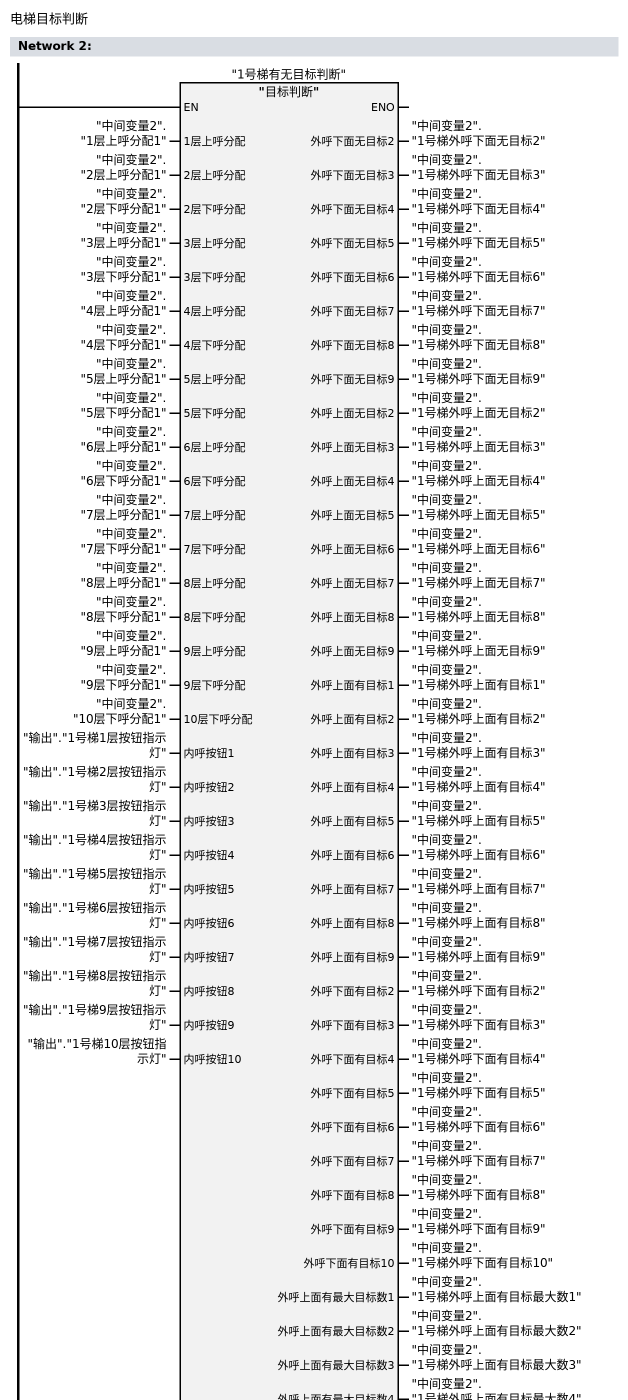
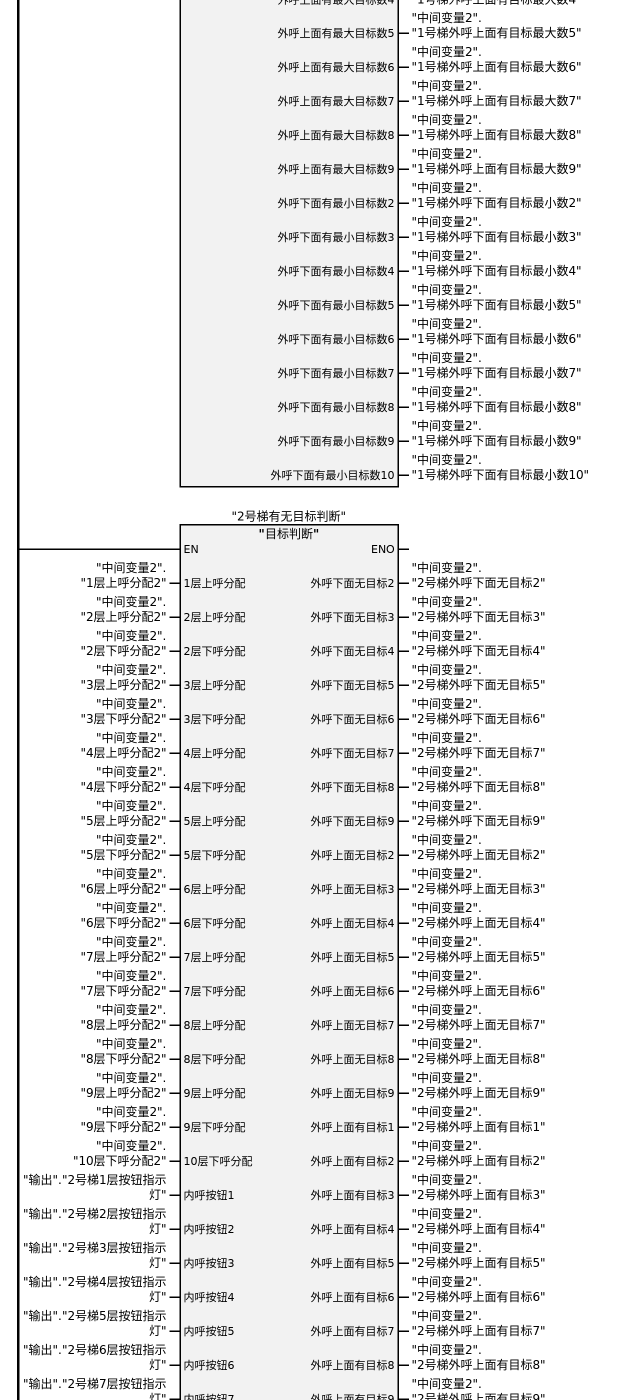
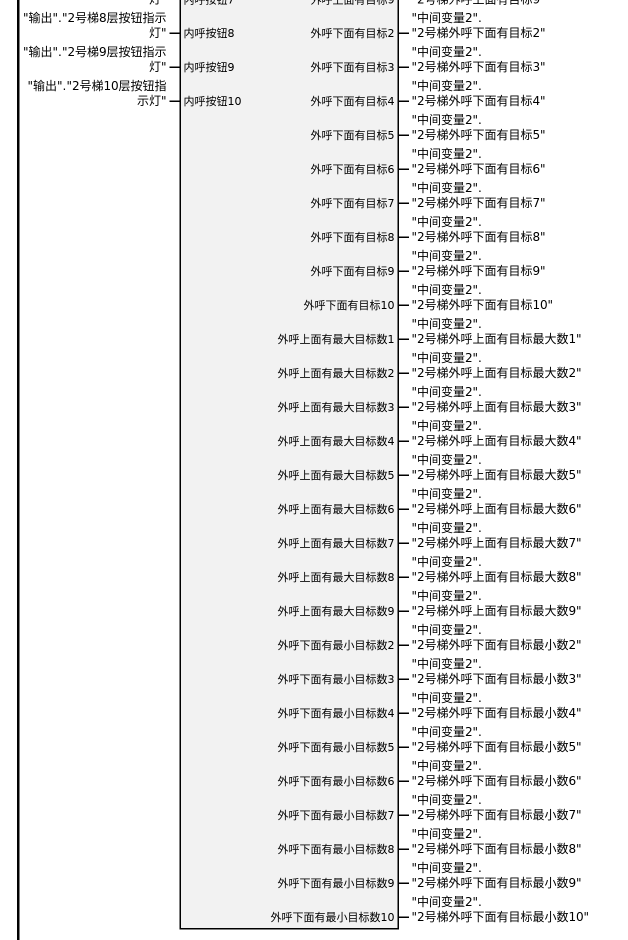
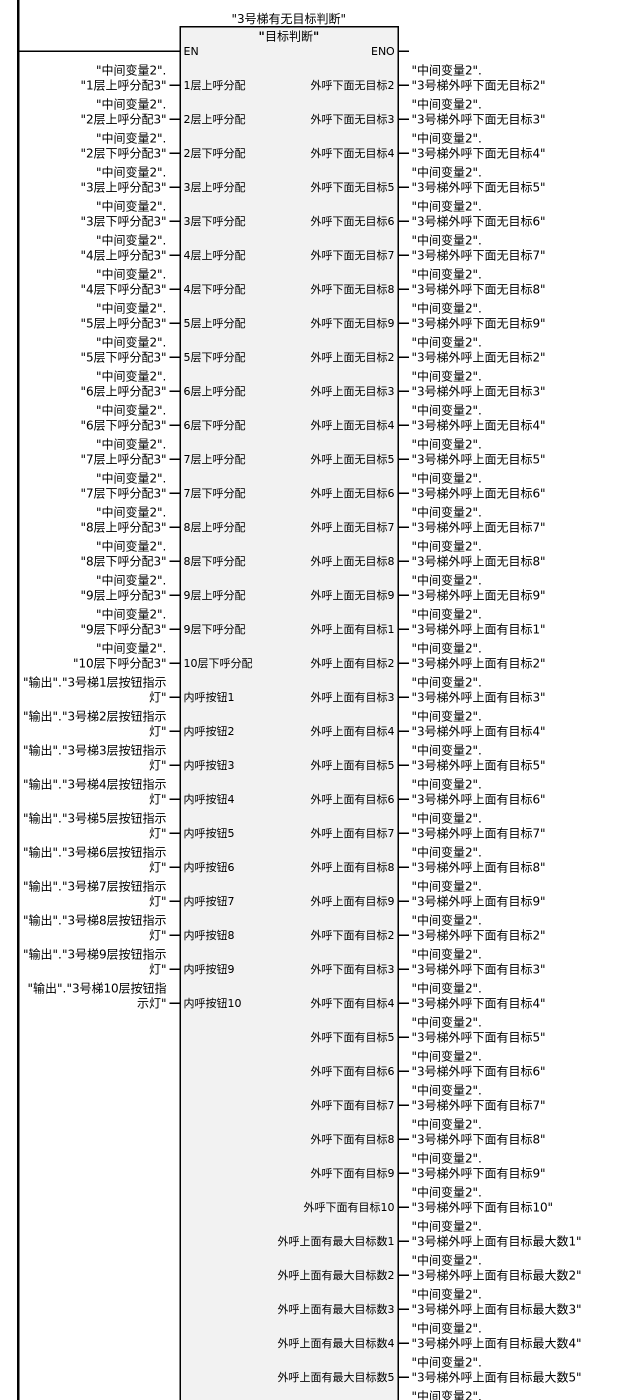
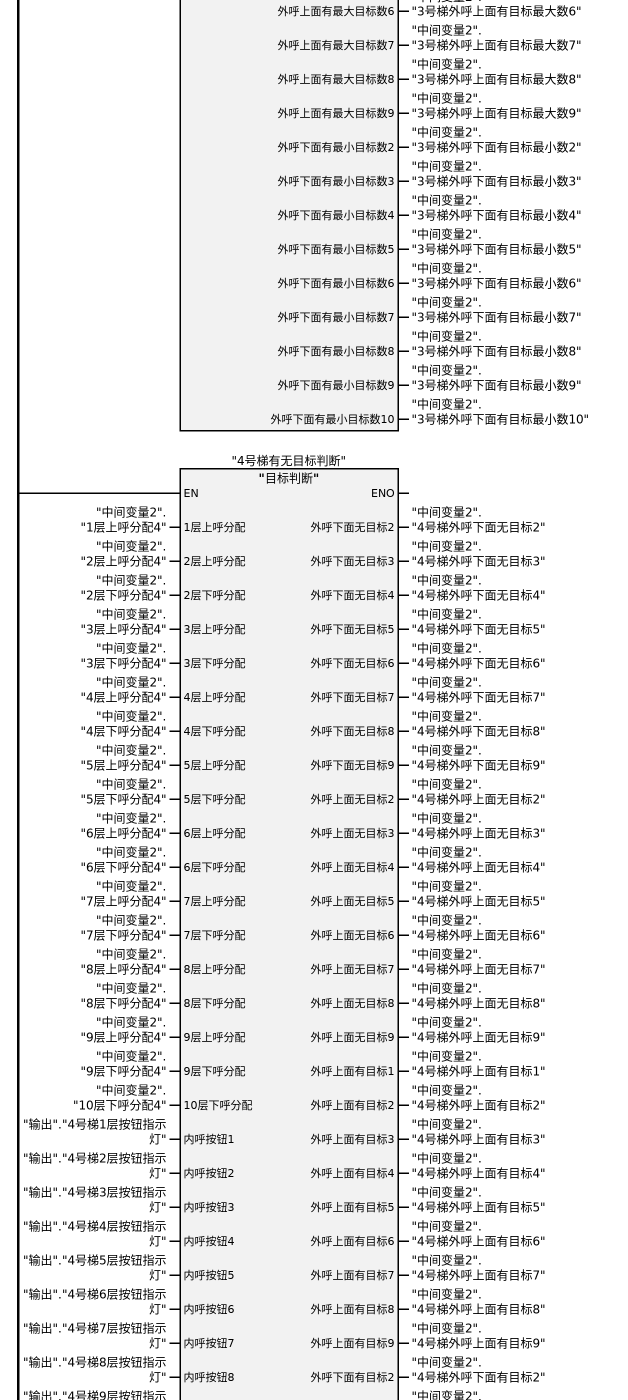
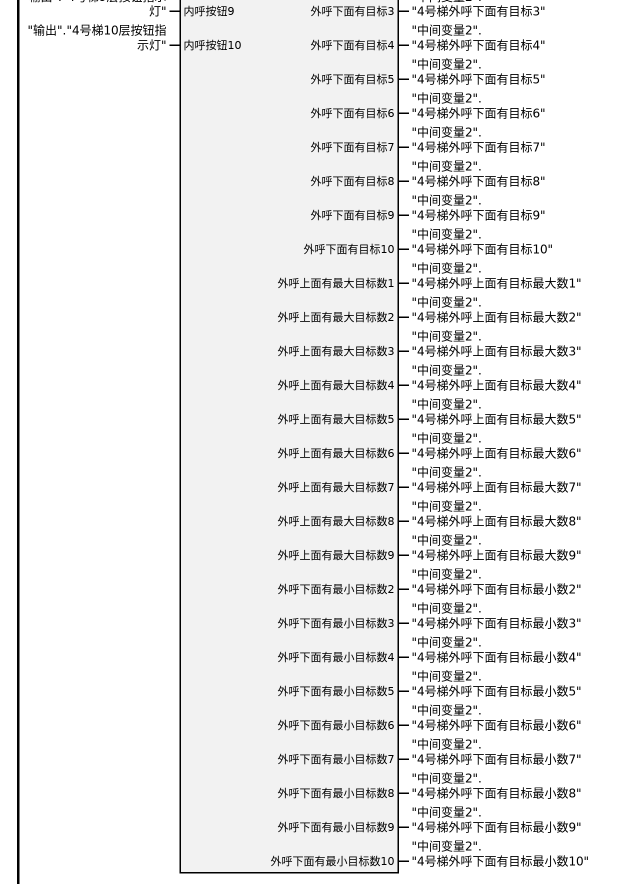
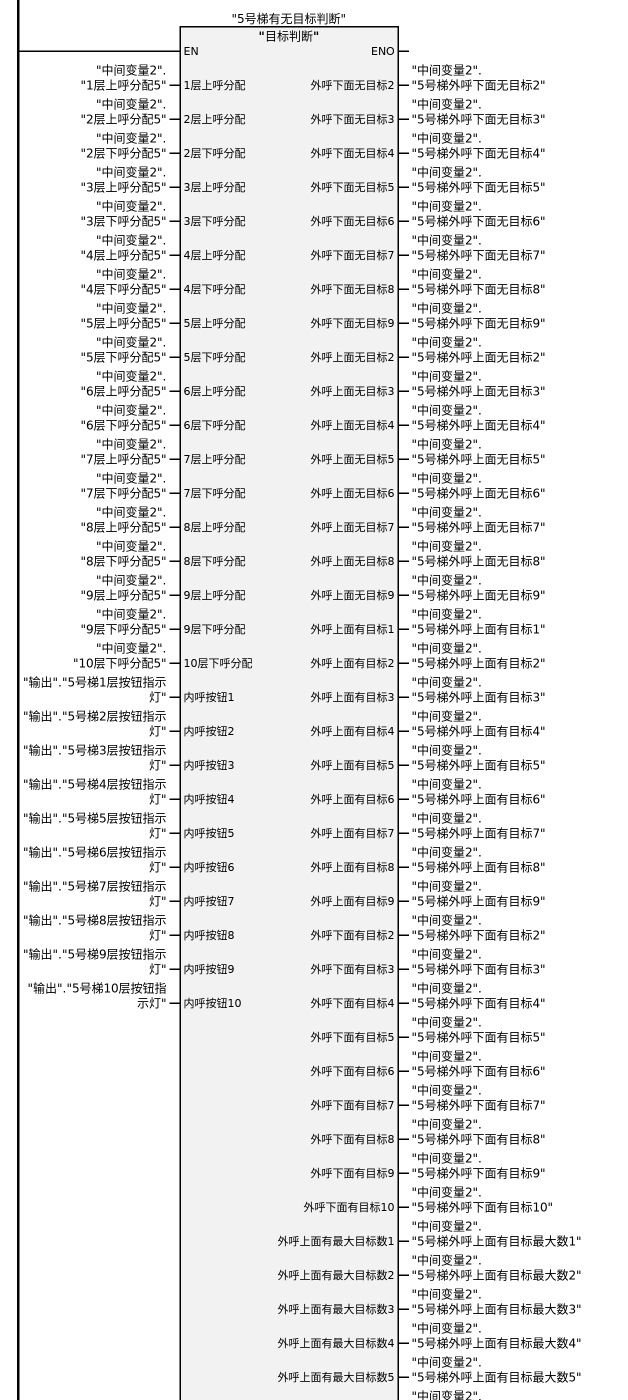
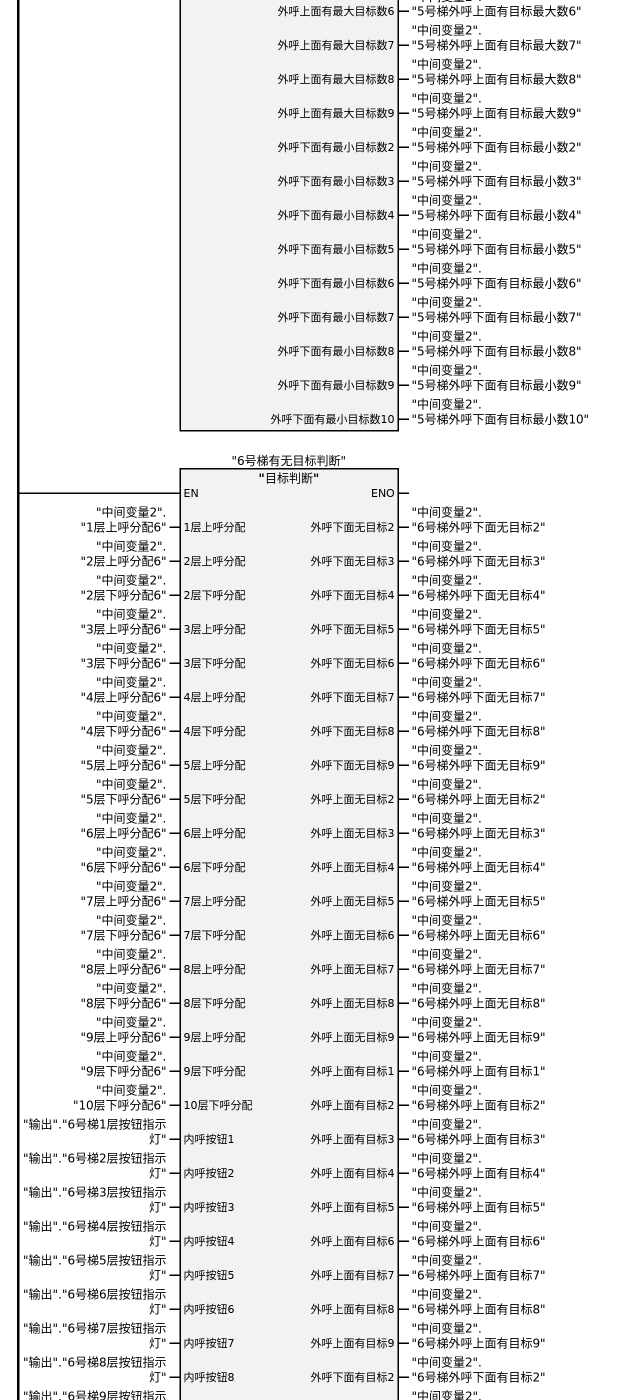
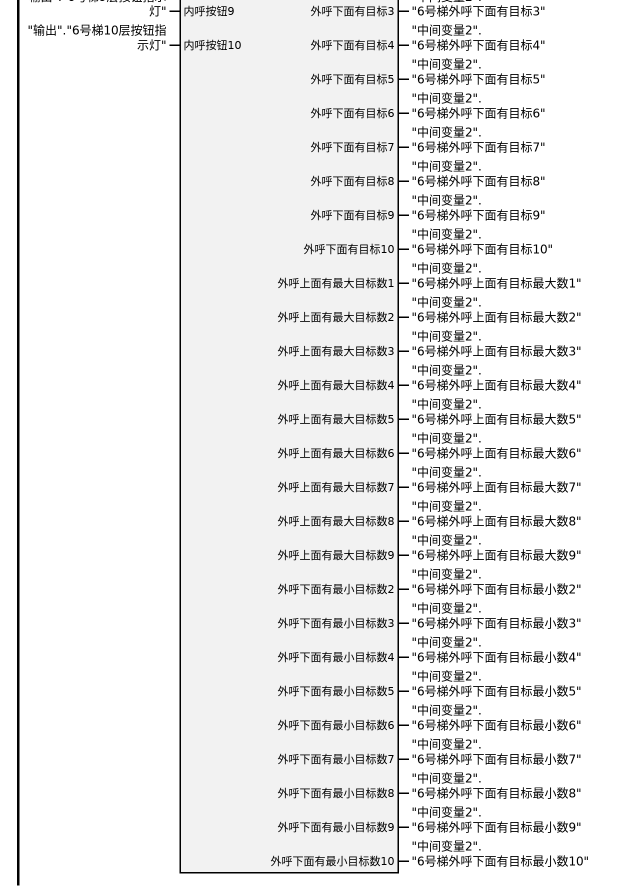
   RUNG wire#powerrail
      "1号梯有无目标判断"("1层上呼分配" := "中间变量2"."1层上呼分配1", "2层上呼分配" := "中间变量2"."2层上呼分配1", "2层下呼分配" := "中间变量2"."2层下呼分配1", "3层上呼分配" := "中间变量2"."3层上呼分配1", "3层下呼分配" := "中间变量2"."3层下呼分配1", "4层上呼分配" := "中间变量2"."4层上呼分配1", "4层下呼分配" := "中间变量2"."4层下呼分配1", "5层上呼分配" := "中间变量2"."5层上呼分配1", "5层下呼分配" := "中间变量2"."5层下呼分配1", "6层上呼分配" := "中间变量2"."6层上呼分配1", "6层下呼分配" := "中间变量2"."6层下呼分配1", "7层上呼分配" := "中间变量2"."7层上呼分配1", "7层下呼分配" := "中间变量2"."7层下呼分配1", "8层上呼分配" := "中间变量2"."8层上呼分配1", "8层下呼分配" := "中间变量2"."8层下呼分配1", "9层上呼分配" := "中间变量2"."9层上呼分配1", "9层下呼分配" := "中间变量2"."9层下呼分配1", "10层下呼分配" := "中间变量2"."10层下呼分配1", 内呼按钮1 := "输出"."1号梯1层按钮指示灯", 内呼按钮2 := "输出"."1号梯2层按钮指示灯", 内呼按钮3 := "输出"."1号梯3层按钮指示灯", 内呼按钮4 := "输出"."1号梯4层按钮指示灯", 内呼按钮5 := "输出"."1号梯5层按钮指示灯", 内呼按钮6 := "输出"."1号梯6层按钮指示灯", 内呼按钮7 := "输出"."1号梯7层按钮指示灯", 内呼按钮8 := "输出"."1号梯8层按钮指示灯", 内呼按钮9 := "输出"."1号梯9层按钮指示灯", 内呼按钮10 := "输出"."1号梯10层按钮指示灯", 外呼下面无目标2 => "中间变量2"."1号梯外呼下面无目标2", 外呼下面无目标3 => "中间变量2"."1号梯外呼下面无目标3", 外呼下面无目标4 => "中间变量2"."1号梯外呼下面无目标4", 外呼下面无目标5 => "中间变量2"."1号梯外呼下面无目标5", 外呼下面无目标6 => "中间变量2"."1号梯外呼下面无目标6", 外呼下面无目标7 => "中间变量2"."1号梯外呼下面无目标7", 外呼下面无目标8 => "中间变量2"."1号梯外呼下面无目标8", 外呼下面无目标9 => "中间变量2"."1号梯外呼下面无目标9", 外呼上面无目标2 => "中间变量2"."1号梯外呼上面无目标2", 外呼上面无目标3 => "中间变量2"."1号梯外呼上面无目标3", 外呼上面无目标4 => "中间变量2"."1号梯外呼上面无目标4", 外呼上面无目标5 => "中间变量2"."1号梯外呼上面无目标5", 外呼上面无目标6 => "中间变量2"."1号梯外呼上面无目标6", 外呼上面无目标7 => "中间变量2"."1号梯外呼上面无目标7", 外呼上面无目标8 => "中间变量2"."1号梯外呼上面无目标8", 外呼上面无目标9 => "中间变量2"."1号梯外呼上面无目标9", 外呼上面有目标1 => "中间变量2"."1号梯外呼上面有目标1", 外呼上面有目标2 => "中间变量2"."1号梯外呼上面有目标2", 外呼上面有目标3 => "中间变量2"."1号梯外呼上面有目标3", 外呼上面有目标4 => "中间变量2"."1号梯外呼上面有目标4", 外呼上面有目标5 => "中间变量2"."1号梯外呼上面有目标5", 外呼上面有目标6 => "中间变量2"."1号梯外呼上面有目标6", 外呼上面有目标7 => "中间变量2"."1号梯外呼上面有目标7", 外呼上面有目标8 => "中间变量2"."1号梯外呼上面有目标8", 外呼上面有目标9 => "中间变量2"."1号梯外呼上面有目标9", 外呼下面有目标2 => "中间变量2"."1号梯外呼下面有目标2", 外呼下面有目标3 => "中间变量2"."1号梯外呼下面有目标3", 外呼下面有目标4 => "中间变量2"."1号梯外呼下面有目标4", 外呼下面有目标5 => "中间变量2"."1号梯外呼下面有目标5", 外呼下面有目标6 => "中间变量2"."1号梯外呼下面有目标6", 外呼下面有目标7 => "中间变量2"."1号梯外呼下面有目标7", 外呼下面有目标8 => "中间变量2"."1号梯外呼下面有目标8", 外呼下面有目标9 => "中间变量2"."1号梯外呼下面有目标9", 外呼下面有目标10 => "中间变量2"."1号梯外呼下面有目标10", 外呼上面有最大目标数1 => "中间变量2"."1号梯外呼上面有目标最大数1", 外呼上面有最大目标数2 => "中间变量2"."1号梯外呼上面有目标最大数2", 外呼上面有最大目标数3 => "中间变量2"."1号梯外呼上面有目标最大数3", 外呼上面有最大目标数4 => "中间变量2"."1号梯外呼上面有目标最大数4", 外呼上面有最大目标数5 => "中间变量2"."1号梯外呼上面有目标最大数5", 外呼上面有最大目标数6 => "中间变量2"."1号梯外呼上面有目标最大数6", 外呼上面有最大目标数7 => "中间变量2"."1号梯外呼上面有目标最大数7", 外呼上面有最大目标数8 => "中间变量2"."1号梯外呼上面有目标最大数8", 外呼上面有最大目标数9 => "中间变量2"."1号梯外呼上面有目标最大数9", 外呼下面有最小目标数2 => "中间变量2"."1号梯外呼下面有目标最小数2", 外呼下面有最小目标数3 => "中间变量2"."1号梯外呼下面有目标最小数3", 外呼下面有最小目标数4 => "中间变量2"."1号梯外呼下面有目标最小数4", 外呼下面有最小目标数5 => "中间变量2"."1号梯外呼下面有目标最小数5", 外呼下面有最小目标数6 => "中间变量2"."1号梯外呼下面有目标最小数6", 外呼下面有最小目标数7 => "中间变量2"."1号梯外呼下面有目标最小数7", 外呼下面有最小目标数8 => "中间变量2"."1号梯外呼下面有目标最小数8", 外呼下面有最小目标数9 => "中间变量2"."1号梯外呼下面有目标最小数9", 外呼下面有最小目标数10 => "中间变量2"."1号梯外呼下面有目标最小数10")
   END_RUNG
   RUNG wire#powerrail
      "2号梯有无目标判断"("1层上呼分配" := "中间变量2"."1层上呼分配2", "2层上呼分配" := "中间变量2"."2层上呼分配2", "2层下呼分配" := "中间变量2"."2层下呼分配2", "3层上呼分配" := "中间变量2"."3层上呼分配2", "3层下呼分配" := "中间变量2"."3层下呼分配2", "4层上呼分配" := "中间变量2"."4层上呼分配2", "4层下呼分配" := "中间变量2"."4层下呼分配2", "5层上呼分配" := "中间变量2"."5层上呼分配2", "5层下呼分配" := "中间变量2"."5层下呼分配2", "6层上呼分配" := "中间变量2"."6层上呼分配2", "6层下呼分配" := "中间变量2"."6层下呼分配2", "7层上呼分配" := "中间变量2"."7层上呼分配2", "7层下呼分配" := "中间变量2"."7层下呼分配2", "8层上呼分配" := "中间变量2"."8层上呼分配2", "8层下呼分配" := "中间变量2"."8层下呼分配2", "9层上呼分配" := "中间变量2"."9层上呼分配2", "9层下呼分配" := "中间变量2"."9层下呼分配2", "10层下呼分配" := "中间变量2"."10层下呼分配2", 内呼按钮1 := "输出"."2号梯1层按钮指示灯", 内呼按钮2 := "输出"."2号梯2层按钮指示灯", 内呼按钮3 := "输出"."2号梯3层按钮指示灯", 内呼按钮4 := "输出"."2号梯4层按钮指示灯", 内呼按钮5 := "输出"."2号梯5层按钮指示灯", 内呼按钮6 := "输出"."2号梯6层按钮指示灯", 内呼按钮7 := "输出"."2号梯7层按钮指示灯", 内呼按钮8 := "输出"."2号梯8层按钮指示灯", 内呼按钮9 := "输出"."2号梯9层按钮指示灯", 内呼按钮10 := "输出"."2号梯10层按钮指示灯", 外呼下面无目标2 => "中间变量2"."2号梯外呼下面无目标2", 外呼下面无目标3 => "中间变量2"."2号梯外呼下面无目标3", 外呼下面无目标4 => "中间变量2"."2号梯外呼下面无目标4", 外呼下面无目标5 => "中间变量2"."2号梯外呼下面无目标5", 外呼下面无目标6 => "中间变量2"."2号梯外呼下面无目标6", 外呼下面无目标7 => "中间变量2"."2号梯外呼下面无目标7", 外呼下面无目标8 => "中间变量2"."2号梯外呼下面无目标8", 外呼下面无目标9 => "中间变量2"."2号梯外呼下面无目标9", 外呼上面无目标2 => "中间变量2"."2号梯外呼上面无目标2", 外呼上面无目标3 => "中间变量2"."2号梯外呼上面无目标3", 外呼上面无目标4 => "中间变量2"."2号梯外呼上面无目标4", 外呼上面无目标5 => "中间变量2"."2号梯外呼上面无目标5", 外呼上面无目标6 => "中间变量2"."2号梯外呼上面无目标6", 外呼上面无目标7 => "中间变量2"."2号梯外呼上面无目标7", 外呼上面无目标8 => "中间变量2"."2号梯外呼上面无目标8", 外呼上面无目标9 => "中间变量2"."2号梯外呼上面无目标9", 外呼上面有目标1 => "中间变量2"."2号梯外呼上面有目标1", 外呼上面有目标2 => "中间变量2"."2号梯外呼上面有目标2", 外呼上面有目标3 => "中间变量2"."2号梯外呼上面有目标3", 外呼上面有目标4 => "中间变量2"."2号梯外呼上面有目标4", 外呼上面有目标5 => "中间变量2"."2号梯外呼上面有目标5", 外呼上面有目标6 => "中间变量2"."2号梯外呼上面有目标6", 外呼上面有目标7 => "中间变量2"."2号梯外呼上面有目标7", 外呼上面有目标8 => "中间变量2"."2号梯外呼上面有目标8", 外呼上面有目标9 => "中间变量2"."2号梯外呼上面有目标9", 外呼下面有目标2 => "中间变量2"."2号梯外呼下面有目标2", 外呼下面有目标3 => "中间变量2"."2号梯外呼下面有目标3", 外呼下面有目标4 => "中间变量2"."2号梯外呼下面有目标4", 外呼下面有目标5 => "中间变量2"."2号梯外呼下面有目标5", 外呼下面有目标6 => "中间变量2"."2号梯外呼下面有目标6", 外呼下面有目标7 => "中间变量2"."2号梯外呼下面有目标7", 外呼下面有目标8 => "中间变量2"."2号梯外呼下面有目标8", 外呼下面有目标9 => "中间变量2"."2号梯外呼下面有目标9", 外呼下面有目标10 => "中间变量2"."2号梯外呼下面有目标10", 外呼上面有最大目标数1 => "中间变量2"."2号梯外呼上面有目标最大数1", 外呼上面有最大目标数2 => "中间变量2"."2号梯外呼上面有目标最大数2", 外呼上面有最大目标数3 => "中间变量2"."2号梯外呼上面有目标最大数3", 外呼上面有最大目标数4 => "中间变量2"."2号梯外呼上面有目标最大数4", 外呼上面有最大目标数5 => "中间变量2"."2号梯外呼上面有目标最大数5", 外呼上面有最大目标数6 => "中间变量2"."2号梯外呼上面有目标最大数6", 外呼上面有最大目标数7 => "中间变量2"."2号梯外呼上面有目标最大数7", 外呼上面有最大目标数8 => "中间变量2"."2号梯外呼上面有目标最大数8", 外呼上面有最大目标数9 => "中间变量2"."2号梯外呼上面有目标最大数9", 外呼下面有最小目标数2 => "中间变量2"."2号梯外呼下面有目标最小数2", 外呼下面有最小目标数3 => "中间变量2"."2号梯外呼下面有目标最小数3", 外呼下面有最小目标数4 => "中间变量2"."2号梯外呼下面有目标最小数4", 外呼下面有最小目标数5 => "中间变量2"."2号梯外呼下面有目标最小数5", 外呼下面有最小目标数6 => "中间变量2"."2号梯外呼下面有目标最小数6", 外呼下面有最小目标数7 => "中间变量2"."2号梯外呼下面有目标最小数7", 外呼下面有最小目标数8 => "中间变量2"."2号梯外呼下面有目标最小数8", 外呼下面有最小目标数9 => "中间变量2"."2号梯外呼下面有目标最小数9", 外呼下面有最小目标数10 => "中间变量2"."2号梯外呼下面有目标最小数10")
   END_RUNG
   RUNG wire#powerrail
      "3号梯有无目标判断"("1层上呼分配" := "中间变量2"."1层上呼分配3", "2层上呼分配" := "中间变量2"."2层上呼分配3", "2层下呼分配" := "中间变量2"."2层下呼分配3", "3层上呼分配" := "中间变量2"."3层上呼分配3", "3层下呼分配" := "中间变量2"."3层下呼分配3", "4层上呼分配" := "中间变量2"."4层上呼分配3", "4层下呼分配" := "中间变量2"."4层下呼分配3", "5层上呼分配" := "中间变量2"."5层上呼分配3", "5层下呼分配" := "中间变量2"."5层下呼分配3", "6层上呼分配" := "中间变量2"."6层上呼分配3", "6层下呼分配" := "中间变量2"."6层下呼分配3", "7层上呼分配" := "中间变量2"."7层上呼分配3", "7层下呼分配" := "中间变量2"."7层下呼分配3", "8层上呼分配" := "中间变量2"."8层上呼分配3", "8层下呼分配" := "中间变量2"."8层下呼分配3", "9层上呼分配" := "中间变量2"."9层上呼分配3", "9层下呼分配" := "中间变量2"."9层下呼分配3", "10层下呼分配" := "中间变量2"."10层下呼分配3", 内呼按钮1 := "输出"."3号梯1层按钮指示灯", 内呼按钮2 := "输出"."3号梯2层按钮指示灯", 内呼按钮3 := "输出"."3号梯3层按钮指示灯", 内呼按钮4 := "输出"."3号梯4层按钮指示灯", 内呼按钮5 := "输出"."3号梯5层按钮指示灯", 内呼按钮6 := "输出"."3号梯6层按钮指示灯", 内呼按钮7 := "输出"."3号梯7层按钮指示灯", 内呼按钮8 := "输出"."3号梯8层按钮指示灯", 内呼按钮9 := "输出"."3号梯9层按钮指示灯", 内呼按钮10 := "输出"."3号梯10层按钮指示灯", 外呼下面无目标2 => "中间变量2"."3号梯外呼下面无目标2", 外呼下面无目标3 => "中间变量2"."3号梯外呼下面无目标3", 外呼下面无目标4 => "中间变量2"."3号梯外呼下面无目标4", 外呼下面无目标5 => "中间变量2"."3号梯外呼下面无目标5", 外呼下面无目标6 => "中间变量2"."3号梯外呼下面无目标6", 外呼下面无目标7 => "中间变量2"."3号梯外呼下面无目标7", 外呼下面无目标8 => "中间变量2"."3号梯外呼下面无目标8", 外呼下面无目标9 => "中间变量2"."3号梯外呼下面无目标9", 外呼上面无目标2 => "中间变量2"."3号梯外呼上面无目标2", 外呼上面无目标3 => "中间变量2"."3号梯外呼上面无目标3", 外呼上面无目标4 => "中间变量2"."3号梯外呼上面无目标4", 外呼上面无目标5 => "中间变量2"."3号梯外呼上面无目标5", 外呼上面无目标6 => "中间变量2"."3号梯外呼上面无目标6", 外呼上面无目标7 => "中间变量2"."3号梯外呼上面无目标7", 外呼上面无目标8 => "中间变量2"."3号梯外呼上面无目标8", 外呼上面无目标9 => "中间变量2"."3号梯外呼上面无目标9", 外呼上面有目标1 => "中间变量2"."3号梯外呼上面有目标1", 外呼上面有目标2 => "中间变量2"."3号梯外呼上面有目标2", 外呼上面有目标3 => "中间变量2"."3号梯外呼上面有目标3", 外呼上面有目标4 => "中间变量2"."3号梯外呼上面有目标4", 外呼上面有目标5 => "中间变量2"."3号梯外呼上面有目标5", 外呼上面有目标6 => "中间变量2"."3号梯外呼上面有目标6", 外呼上面有目标7 => "中间变量2"."3号梯外呼上面有目标7", 外呼上面有目标8 => "中间变量2"."3号梯外呼上面有目标8", 外呼上面有目标9 => "中间变量2"."3号梯外呼上面有目标9", 外呼下面有目标2 => "中间变量2"."3号梯外呼下面有目标2", 外呼下面有目标3 => "中间变量2"."3号梯外呼下面有目标3", 外呼下面有目标4 => "中间变量2"."3号梯外呼下面有目标4", 外呼下面有目标5 => "中间变量2"."3号梯外呼下面有目标5", 外呼下面有目标6 => "中间变量2"."3号梯外呼下面有目标6", 外呼下面有目标7 => "中间变量2"."3号梯外呼下面有目标7", 外呼下面有目标8 => "中间变量2"."3号梯外呼下面有目标8", 外呼下面有目标9 => "中间变量2"."3号梯外呼下面有目标9", 外呼下面有目标10 => "中间变量2"."3号梯外呼下面有目标10", 外呼上面有最大目标数1 => "中间变量2"."3号梯外呼上面有目标最大数1", 外呼上面有最大目标数2 => "中间变量2"."3号梯外呼上面有目标最大数2", 外呼上面有最大目标数3 => "中间变量2"."3号梯外呼上面有目标最大数3", 外呼上面有最大目标数4 => "中间变量2"."3号梯外呼上面有目标最大数4", 外呼上面有最大目标数5 => "中间变量2"."3号梯外呼上面有目标最大数5", 外呼上面有最大目标数6 => "中间变量2"."3号梯外呼上面有目标最大数6", 外呼上面有最大目标数7 => "中间变量2"."3号梯外呼上面有目标最大数7", 外呼上面有最大目标数8 => "中间变量2"."3号梯外呼上面有目标最大数8", 外呼上面有最大目标数9 => "中间变量2"."3号梯外呼上面有目标最大数9", 外呼下面有最小目标数2 => "中间变量2"."3号梯外呼下面有目标最小数2", 外呼下面有最小目标数3 => "中间变量2"."3号梯外呼下面有目标最小数3", 外呼下面有最小目标数4 => "中间变量2"."3号梯外呼下面有目标最小数4", 外呼下面有最小目标数5 => "中间变量2"."3号梯外呼下面有目标最小数5", 外呼下面有最小目标数6 => "中间变量2"."3号梯外呼下面有目标最小数6", 外呼下面有最小目标数7 => "中间变量2"."3号梯外呼下面有目标最小数7", 外呼下面有最小目标数8 => "中间变量2"."3号梯外呼下面有目标最小数8", 外呼下面有最小目标数9 => "中间变量2"."3号梯外呼下面有目标最小数9", 外呼下面有最小目标数10 => "中间变量2"."3号梯外呼下面有目标最小数10")
   END_RUNG
   RUNG wire#powerrail
      "4号梯有无目标判断"("1层上呼分配" := "中间变量2"."1层上呼分配4", "2层上呼分配" := "中间变量2"."2层上呼分配4", "2层下呼分配" := "中间变量2"."2层下呼分配4", "3层上呼分配" := "中间变量2"."3层上呼分配4", "3层下呼分配" := "中间变量2"."3层下呼分配4", "4层上呼分配" := "中间变量2"."4层上呼分配4", "4层下呼分配" := "中间变量2"."4层下呼分配4", "5层上呼分配" := "中间变量2"."5层上呼分配4", "5层下呼分配" := "中间变量2"."5层下呼分配4", "6层上呼分配" := "中间变量2"."6层上呼分配4", "6层下呼分配" := "中间变量2"."6层下呼分配4", "7层上呼分配" := "中间变量2"."7层上呼分配4", "7层下呼分配" := "中间变量2"."7层下呼分配4", "8层上呼分配" := "中间变量2"."8层上呼分配4", "8层下呼分配" := "中间变量2"."8层下呼分配4", "9层上呼分配" := "中间变量2"."9层上呼分配4", "9层下呼分配" := "中间变量2"."9层下呼分配4", "10层下呼分配" := "中间变量2"."10层下呼分配4", 内呼按钮1 := "输出"."4号梯1层按钮指示灯", 内呼按钮2 := "输出"."4号梯2层按钮指示灯", 内呼按钮3 := "输出"."4号梯3层按钮指示灯", 内呼按钮4 := "输出"."4号梯4层按钮指示灯", 内呼按钮5 := "输出"."4号梯5层按钮指示灯", 内呼按钮6 := "输出"."4号梯6层按钮指示灯", 内呼按钮7 := "输出"."4号梯7层按钮指示灯", 内呼按钮8 := "输出"."4号梯8层按钮指示灯", 内呼按钮9 := "输出"."4号梯9层按钮指示灯", 内呼按钮10 := "输出"."4号梯10层按钮指示灯", 外呼下面无目标2 => "中间变量2"."4号梯外呼下面无目标2", 外呼下面无目标3 => "中间变量2"."4号梯外呼下面无目标3", 外呼下面无目标4 => "中间变量2"."4号梯外呼下面无目标4", 外呼下面无目标5 => "中间变量2"."4号梯外呼下面无目标5", 外呼下面无目标6 => "中间变量2"."4号梯外呼下面无目标6", 外呼下面无目标7 => "中间变量2"."4号梯外呼下面无目标7", 外呼下面无目标8 => "中间变量2"."4号梯外呼下面无目标8", 外呼下面无目标9 => "中间变量2"."4号梯外呼下面无目标9", 外呼上面无目标2 => "中间变量2"."4号梯外呼上面无目标2", 外呼上面无目标3 => "中间变量2"."4号梯外呼上面无目标3", 外呼上面无目标4 => "中间变量2"."4号梯外呼上面无目标4", 外呼上面无目标5 => "中间变量2"."4号梯外呼上面无目标5", 外呼上面无目标6 => "中间变量2"."4号梯外呼上面无目标6", 外呼上面无目标7 => "中间变量2"."4号梯外呼上面无目标7", 外呼上面无目标8 => "中间变量2"."4号梯外呼上面无目标8", 外呼上面无目标9 => "中间变量2"."4号梯外呼上面无目标9", 外呼上面有目标1 => "中间变量2"."4号梯外呼上面有目标1", 外呼上面有目标2 => "中间变量2"."4号梯外呼上面有目标2", 外呼上面有目标3 => "中间变量2"."4号梯外呼上面有目标3", 外呼上面有目标4 => "中间变量2"."4号梯外呼上面有目标4", 外呼上面有目标5 => "中间变量2"."4号梯外呼上面有目标5", 外呼上面有目标6 => "中间变量2"."4号梯外呼上面有目标6", 外呼上面有目标7 => "中间变量2"."4号梯外呼上面有目标7", 外呼上面有目标8 => "中间变量2"."4号梯外呼上面有目标8", 外呼上面有目标9 => "中间变量2"."4号梯外呼上面有目标9", 外呼下面有目标2 => "中间变量2"."4号梯外呼下面有目标2", 外呼下面有目标3 => "中间变量2"."4号梯外呼下面有目标3", 外呼下面有目标4 => "中间变量2"."4号梯外呼下面有目标4", 外呼下面有目标5 => "中间变量2"."4号梯外呼下面有目标5", 外呼下面有目标6 => "中间变量2"."4号梯外呼下面有目标6", 外呼下面有目标7 => "中间变量2"."4号梯外呼下面有目标7", 外呼下面有目标8 => "中间变量2"."4号梯外呼下面有目标8", 外呼下面有目标9 => "中间变量2"."4号梯外呼下面有目标9", 外呼下面有目标10 => "中间变量2"."4号梯外呼下面有目标10", 外呼上面有最大目标数1 => "中间变量2"."4号梯外呼上面有目标最大数1", 外呼上面有最大目标数2 => "中间变量2"."4号梯外呼上面有目标最大数2", 外呼上面有最大目标数3 => "中间变量2"."4号梯外呼上面有目标最大数3", 外呼上面有最大目标数4 => "中间变量2"."4号梯外呼上面有目标最大数4", 外呼上面有最大目标数5 => "中间变量2"."4号梯外呼上面有目标最大数5", 外呼上面有最大目标数6 => "中间变量2"."4号梯外呼上面有目标最大数6", 外呼上面有最大目标数7 => "中间变量2"."4号梯外呼上面有目标最大数7", 外呼上面有最大目标数8 => "中间变量2"."4号梯外呼上面有目标最大数8", 外呼上面有最大目标数9 => "中间变量2"."4号梯外呼上面有目标最大数9", 外呼下面有最小目标数2 => "中间变量2"."4号梯外呼下面有目标最小数2", 外呼下面有最小目标数3 => "中间变量2"."4号梯外呼下面有目标最小数3", 外呼下面有最小目标数4 => "中间变量2"."4号梯外呼下面有目标最小数4", 外呼下面有最小目标数5 => "中间变量2"."4号梯外呼下面有目标最小数5", 外呼下面有最小目标数6 => "中间变量2"."4号梯外呼下面有目标最小数6", 外呼下面有最小目标数7 => "中间变量2"."4号梯外呼下面有目标最小数7", 外呼下面有最小目标数8 => "中间变量2"."4号梯外呼下面有目标最小数8", 外呼下面有最小目标数9 => "中间变量2"."4号梯外呼下面有目标最小数9", 外呼下面有最小目标数10 => "中间变量2"."4号梯外呼下面有目标最小数10")
   END_RUNG
   RUNG wire#powerrail
      "5号梯有无目标判断"("1层上呼分配" := "中间变量2"."1层上呼分配5", "2层上呼分配" := "中间变量2"."2层上呼分配5", "2层下呼分配" := "中间变量2"."2层下呼分配5", "3层上呼分配" := "中间变量2"."3层上呼分配5", "3层下呼分配" := "中间变量2"."3层下呼分配5", "4层上呼分配" := "中间变量2"."4层上呼分配5", "4层下呼分配" := "中间变量2"."4层下呼分配5", "5层上呼分配" := "中间变量2"."5层上呼分配5", "5层下呼分配" := "中间变量2"."5层下呼分配5", "6层上呼分配" := "中间变量2"."6层上呼分配5", "6层下呼分配" := "中间变量2"."6层下呼分配5", "7层上呼分配" := "中间变量2"."7层上呼分配5", "7层下呼分配" := "中间变量2"."7层下呼分配5", "8层上呼分配" := "中间变量2"."8层上呼分配5", "8层下呼分配" := "中间变量2"."8层下呼分配5", "9层上呼分配" := "中间变量2"."9层上呼分配5", "9层下呼分配" := "中间变量2"."9层下呼分配5", "10层下呼分配" := "中间变量2"."10层下呼分配5", 内呼按钮1 := "输出"."5号梯1层按钮指示灯", 内呼按钮2 := "输出"."5号梯2层按钮指示灯", 内呼按钮3 := "输出"."5号梯3层按钮指示灯", 内呼按钮4 := "输出"."5号梯4层按钮指示灯", 内呼按钮5 := "输出"."5号梯5层按钮指示灯", 内呼按钮6 := "输出"."5号梯6层按钮指示灯", 内呼按钮7 := "输出"."5号梯7层按钮指示灯", 内呼按钮8 := "输出"."5号梯8层按钮指示灯", 内呼按钮9 := "输出"."5号梯9层按钮指示灯", 内呼按钮10 := "输出"."5号梯10层按钮指示灯", 外呼下面无目标2 => "中间变量2"."5号梯外呼下面无目标2", 外呼下面无目标3 => "中间变量2"."5号梯外呼下面无目标3", 外呼下面无目标4 => "中间变量2"."5号梯外呼下面无目标4", 外呼下面无目标5 => "中间变量2"."5号梯外呼下面无目标5", 外呼下面无目标6 => "中间变量2"."5号梯外呼下面无目标6", 外呼下面无目标7 => "中间变量2"."5号梯外呼下面无目标7", 外呼下面无目标8 => "中间变量2"."5号梯外呼下面无目标8", 外呼下面无目标9 => "中间变量2"."5号梯外呼下面无目标9", 外呼上面无目标2 => "中间变量2"."5号梯外呼上面无目标2", 外呼上面无目标3 => "中间变量2"."5号梯外呼上面无目标3", 外呼上面无目标4 => "中间变量2"."5号梯外呼上面无目标4", 外呼上面无目标5 => "中间变量2"."5号梯外呼上面无目标5", 外呼上面无目标6 => "中间变量2"."5号梯外呼上面无目标6", 外呼上面无目标7 => "中间变量2"."5号梯外呼上面无目标7", 外呼上面无目标8 => "中间变量2"."5号梯外呼上面无目标8", 外呼上面无目标9 => "中间变量2"."5号梯外呼上面无目标9", 外呼上面有目标1 => "中间变量2"."5号梯外呼上面有目标1", 外呼上面有目标2 => "中间变量2"."5号梯外呼上面有目标2", 外呼上面有目标3 => "中间变量2"."5号梯外呼上面有目标3", 外呼上面有目标4 => "中间变量2"."5号梯外呼上面有目标4", 外呼上面有目标5 => "中间变量2"."5号梯外呼上面有目标5", 外呼上面有目标6 => "中间变量2"."5号梯外呼上面有目标6", 外呼上面有目标7 => "中间变量2"."5号梯外呼上面有目标7", 外呼上面有目标8 => "中间变量2"."5号梯外呼上面有目标8", 外呼上面有目标9 => "中间变量2"."5号梯外呼上面有目标9", 外呼下面有目标2 => "中间变量2"."5号梯外呼下面有目标2", 外呼下面有目标3 => "中间变量2"."5号梯外呼下面有目标3", 外呼下面有目标4 => "中间变量2"."5号梯外呼下面有目标4", 外呼下面有目标5 => "中间变量2"."5号梯外呼下面有目标5", 外呼下面有目标6 => "中间变量2"."5号梯外呼下面有目标6", 外呼下面有目标7 => "中间变量2"."5号梯外呼下面有目标7", 外呼下面有目标8 => "中间变量2"."5号梯外呼下面有目标8", 外呼下面有目标9 => "中间变量2"."5号梯外呼下面有目标9", 外呼下面有目标10 => "中间变量2"."5号梯外呼下面有目标10", 外呼上面有最大目标数1 => "中间变量2"."5号梯外呼上面有目标最大数1", 外呼上面有最大目标数2 => "中间变量2"."5号梯外呼上面有目标最大数2", 外呼上面有最大目标数3 => "中间变量2"."5号梯外呼上面有目标最大数3", 外呼上面有最大目标数4 => "中间变量2"."5号梯外呼上面有目标最大数4", 外呼上面有最大目标数5 => "中间变量2"."5号梯外呼上面有目标最大数5", 外呼上面有最大目标数6 => "中间变量2"."5号梯外呼上面有目标最大数6", 外呼上面有最大目标数7 => "中间变量2"."5号梯外呼上面有目标最大数7", 外呼上面有最大目标数8 => "中间变量2"."5号梯外呼上面有目标最大数8", 外呼上面有最大目标数9 => "中间变量2"."5号梯外呼上面有目标最大数9", 外呼下面有最小目标数2 => "中间变量2"."5号梯外呼下面有目标最小数2", 外呼下面有最小目标数3 => "中间变量2"."5号梯外呼下面有目标最小数3", 外呼下面有最小目标数4 => "中间变量2"."5号梯外呼下面有目标最小数4", 外呼下面有最小目标数5 => "中间变量2"."5号梯外呼下面有目标最小数5", 外呼下面有最小目标数6 => "中间变量2"."5号梯外呼下面有目标最小数6", 外呼下面有最小目标数7 => "中间变量2"."5号梯外呼下面有目标最小数7", 外呼下面有最小目标数8 => "中间变量2"."5号梯外呼下面有目标最小数8", 外呼下面有最小目标数9 => "中间变量2"."5号梯外呼下面有目标最小数9", 外呼下面有最小目标数10 => "中间变量2"."5号梯外呼下面有目标最小数10")
   END_RUNG
   RUNG wire#powerrail
      "6号梯有无目标判断"("1层上呼分配" := "中间变量2"."1层上呼分配6", "2层上呼分配" := "中间变量2"."2层上呼分配6", "2层下呼分配" := "中间变量2"."2层下呼分配6", "3层上呼分配" := "中间变量2"."3层上呼分配6", "3层下呼分配" := "中间变量2"."3层下呼分配6", "4层上呼分配" := "中间变量2"."4层上呼分配6", "4层下呼分配" := "中间变量2"."4层下呼分配6", "5层上呼分配" := "中间变量2"."5层上呼分配6", "5层下呼分配" := "中间变量2"."5层下呼分配6", "6层上呼分配" := "中间变量2"."6层上呼分配6", "6层下呼分配" := "中间变量2"."6层下呼分配6", "7层上呼分配" := "中间变量2"."7层上呼分配6", "7层下呼分配" := "中间变量2"."7层下呼分配6", "8层上呼分配" := "中间变量2"."8层上呼分配6", "8层下呼分配" := "中间变量2"."8层下呼分配6", "9层上呼分配" := "中间变量2"."9层上呼分配6", "9层下呼分配" := "中间变量2"."9层下呼分配6", "10层下呼分配" := "中间变量2"."10层下呼分配6", 内呼按钮1 := "输出"."6号梯1层按钮指示灯", 内呼按钮2 := "输出"."6号梯2层按钮指示灯", 内呼按钮3 := "输出"."6号梯3层按钮指示灯", 内呼按钮4 := "输出"."6号梯4层按钮指示灯", 内呼按钮5 := "输出"."6号梯5层按钮指示灯", 内呼按钮6 := "输出"."6号梯6层按钮指示灯", 内呼按钮7 := "输出"."6号梯7层按钮指示灯", 内呼按钮8 := "输出"."6号梯8层按钮指示灯", 内呼按钮9 := "输出"."6号梯9层按钮指示灯", 内呼按钮10 := "输出"."6号梯10层按钮指示灯", 外呼下面无目标2 => "中间变量2"."6号梯外呼下面无目标2", 外呼下面无目标3 => "中间变量2"."6号梯外呼下面无目标3", 外呼下面无目标4 => "中间变量2"."6号梯外呼下面无目标4", 外呼下面无目标5 => "中间变量2"."6号梯外呼下面无目标5", 外呼下面无目标6 => "中间变量2"."6号梯外呼下面无目标6", 外呼下面无目标7 => "中间变量2"."6号梯外呼下面无目标7", 外呼下面无目标8 => "中间变量2"."6号梯外呼下面无目标8", 外呼下面无目标9 => "中间变量2"."6号梯外呼下面无目标9", 外呼上面无目标2 => "中间变量2"."6号梯外呼上面无目标2", 外呼上面无目标3 => "中间变量2"."6号梯外呼上面无目标3", 外呼上面无目标4 => "中间变量2"."6号梯外呼上面无目标4", 外呼上面无目标5 => "中间变量2"."6号梯外呼上面无目标5", 外呼上面无目标6 => "中间变量2"."6号梯外呼上面无目标6", 外呼上面无目标7 => "中间变量2"."6号梯外呼上面无目标7", 外呼上面无目标8 => "中间变量2"."6号梯外呼上面无目标8", 外呼上面无目标9 => "中间变量2"."6号梯外呼上面无目标9", 外呼上面有目标1 => "中间变量2"."6号梯外呼上面有目标1", 外呼上面有目标2 => "中间变量2"."6号梯外呼上面有目标2", 外呼上面有目标3 => "中间变量2"."6号梯外呼上面有目标3", 外呼上面有目标4 => "中间变量2"."6号梯外呼上面有目标4", 外呼上面有目标5 => "中间变量2"."6号梯外呼上面有目标5", 外呼上面有目标6 => "中间变量2"."6号梯外呼上面有目标6", 外呼上面有目标7 => "中间变量2"."6号梯外呼上面有目标7", 外呼上面有目标8 => "中间变量2"."6号梯外呼上面有目标8", 外呼上面有目标9 => "中间变量2"."6号梯外呼上面有目标9", 外呼下面有目标2 => "中间变量2"."6号梯外呼下面有目标2", 外呼下面有目标3 => "中间变量2"."6号梯外呼下面有目标3", 外呼下面有目标4 => "中间变量2"."6号梯外呼下面有目标4", 外呼下面有目标5 => "中间变量2"."6号梯外呼下面有目标5", 外呼下面有目标6 => "中间变量2"."6号梯外呼下面有目标6", 外呼下面有目标7 => "中间变量2"."6号梯外呼下面有目标7", 外呼下面有目标8 => "中间变量2"."6号梯外呼下面有目标8", 外呼下面有目标9 => "中间变量2"."6号梯外呼下面有目标9", 外呼下面有目标10 => "中间变量2"."6号梯外呼下面有目标10", 外呼上面有最大目标数1 => "中间变量2"."6号梯外呼上面有目标最大数1", 外呼上面有最大目标数2 => "中间变量2"."6号梯外呼上面有目标最大数2", 外呼上面有最大目标数3 => "中间变量2"."6号梯外呼上面有目标最大数3", 外呼上面有最大目标数4 => "中间变量2"."6号梯外呼上面有目标最大数4", 外呼上面有最大目标数5 => "中间变量2"."6号梯外呼上面有目标最大数5", 外呼上面有最大目标数6 => "中间变量2"."6号梯外呼上面有目标最大数6", 外呼上面有最大目标数7 => "中间变量2"."6号梯外呼上面有目标最大数7", 外呼上面有最大目标数8 => "中间变量2"."6号梯外呼上面有目标最大数8", 外呼上面有最大目标数9 => "中间变量2"."6号梯外呼上面有目标最大数9", 外呼下面有最小目标数2 => "中间变量2"."6号梯外呼下面有目标最小数2", 外呼下面有最小目标数3 => "中间变量2"."6号梯外呼下面有目标最小数3", 外呼下面有最小目标数4 => "中间变量2"."6号梯外呼下面有目标最小数4", 外呼下面有最小目标数5 => "中间变量2"."6号梯外呼下面有目标最小数5", 外呼下面有最小目标数6 => "中间变量2"."6号梯外呼下面有目标最小数6", 外呼下面有最小目标数7 => "中间变量2"."6号梯外呼下面有目标最小数7", 外呼下面有最小目标数8 => "中间变量2"."6号梯外呼下面有目标最小数8", 外呼下面有最小目标数9 => "中间变量2"."6号梯外呼下面有目标最小数9", 外呼下面有最小目标数10 => "中间变量2"."6号梯外呼下面有目标最小数10")
   END_RUNG
   // the same network as SCL:
   "1号梯有无目标判断"("1层上呼分配" := "中间变量2"."1层上呼分配1",   // "目标判断"
               "2层上呼分配" := "中间变量2"."2层上呼分配1",
               "2层下呼分配" := "中间变量2"."2层下呼分配1",
               "3层上呼分配" := "中间变量2"."3层上呼分配1",
               "3层下呼分配" := "中间变量2"."3层下呼分配1",
               "4层上呼分配" := "中间变量2"."4层上呼分配1",
               "4层下呼分配" := "中间变量2"."4层下呼分配1",
               "5层上呼分配" := "中间变量2"."5层上呼分配1",
               "5层下呼分配" := "中间变量2"."5层下呼分配1",
               "6层上呼分配" := "中间变量2"."6层上呼分配1",
               "6层下呼分配" := "中间变量2"."6层下呼分配1",
               "7层上呼分配" := "中间变量2"."7层上呼分配1",
               "7层下呼分配" := "中间变量2"."7层下呼分配1",
               "8层上呼分配" := "中间变量2"."8层上呼分配1",
               "8层下呼分配" := "中间变量2"."8层下呼分配1",
               "9层上呼分配" := "中间变量2"."9层上呼分配1",
               "9层下呼分配" := "中间变量2"."9层下呼分配1",
               "10层下呼分配" := "中间变量2"."10层下呼分配1",
               内呼按钮1 := "输出"."1号梯1层按钮指示灯",
               内呼按钮2 := "输出"."1号梯2层按钮指示灯",
               内呼按钮3 := "输出"."1号梯3层按钮指示灯",
               内呼按钮4 := "输出"."1号梯4层按钮指示灯",
               内呼按钮5 := "输出"."1号梯5层按钮指示灯",
               内呼按钮6 := "输出"."1号梯6层按钮指示灯",
               内呼按钮7 := "输出"."1号梯7层按钮指示灯",
               内呼按钮8 := "输出"."1号梯8层按钮指示灯",
               内呼按钮9 := "输出"."1号梯9层按钮指示灯",
               内呼按钮10 := "输出"."1号梯10层按钮指示灯",
               外呼下面无目标2 => "中间变量2"."1号梯外呼下面无目标2",
               外呼下面无目标3 => "中间变量2"."1号梯外呼下面无目标3",
               外呼下面无目标4 => "中间变量2"."1号梯外呼下面无目标4",
               外呼下面无目标5 => "中间变量2"."1号梯外呼下面无目标5",
               外呼下面无目标6 => "中间变量2"."1号梯外呼下面无目标6",
               外呼下面无目标7 => "中间变量2"."1号梯外呼下面无目标7",
               外呼下面无目标8 => "中间变量2"."1号梯外呼下面无目标8",
               外呼下面无目标9 => "中间变量2"."1号梯外呼下面无目标9",
               外呼上面无目标2 => "中间变量2"."1号梯外呼上面无目标2",
               外呼上面无目标3 => "中间变量2"."1号梯外呼上面无目标3",
               外呼上面无目标4 => "中间变量2"."1号梯外呼上面无目标4",
               外呼上面无目标5 => "中间变量2"."1号梯外呼上面无目标5",
               外呼上面无目标6 => "中间变量2"."1号梯外呼上面无目标6",
               外呼上面无目标7 => "中间变量2"."1号梯外呼上面无目标7",
               外呼上面无目标8 => "中间变量2"."1号梯外呼上面无目标8",
               外呼上面无目标9 => "中间变量2"."1号梯外呼上面无目标9",
               外呼上面有目标1 => "中间变量2"."1号梯外呼上面有目标1",
               外呼上面有目标2 => "中间变量2"."1号梯外呼上面有目标2",
               外呼上面有目标3 => "中间变量2"."1号梯外呼上面有目标3",
               外呼上面有目标4 => "中间变量2"."1号梯外呼上面有目标4",
               外呼上面有目标5 => "中间变量2"."1号梯外呼上面有目标5",
               外呼上面有目标6 => "中间变量2"."1号梯外呼上面有目标6",
               外呼上面有目标7 => "中间变量2"."1号梯外呼上面有目标7",
               外呼上面有目标8 => "中间变量2"."1号梯外呼上面有目标8",
               外呼上面有目标9 => "中间变量2"."1号梯外呼上面有目标9",
               外呼下面有目标2 => "中间变量2"."1号梯外呼下面有目标2",
               外呼下面有目标3 => "中间变量2"."1号梯外呼下面有目标3",
               外呼下面有目标4 => "中间变量2"."1号梯外呼下面有目标4",
               外呼下面有目标5 => "中间变量2"."1号梯外呼下面有目标5",
               外呼下面有目标6 => "中间变量2"."1号梯外呼下面有目标6",
               外呼下面有目标7 => "中间变量2"."1号梯外呼下面有目标7",
               外呼下面有目标8 => "中间变量2"."1号梯外呼下面有目标8",
               外呼下面有目标9 => "中间变量2"."1号梯外呼下面有目标9",
               外呼下面有目标10 => "中间变量2"."1号梯外呼下面有目标10",
               外呼上面有最大目标数1 => "中间变量2"."1号梯外呼上面有目标最大数1",
               外呼上面有最大目标数2 => "中间变量2"."1号梯外呼上面有目标最大数2",
               外呼上面有最大目标数3 => "中间变量2"."1号梯外呼上面有目标最大数3",
               外呼上面有最大目标数4 => "中间变量2"."1号梯外呼上面有目标最大数4",
               外呼上面有最大目标数5 => "中间变量2"."1号梯外呼上面有目标最大数5",
               外呼上面有最大目标数6 => "中间变量2"."1号梯外呼上面有目标最大数6",
               外呼上面有最大目标数7 => "中间变量2"."1号梯外呼上面有目标最大数7",
               外呼上面有最大目标数8 => "中间变量2"."1号梯外呼上面有目标最大数8",
               外呼上面有最大目标数9 => "中间变量2"."1号梯外呼上面有目标最大数9",
               外呼下面有最小目标数2 => "中间变量2"."1号梯外呼下面有目标最小数2",
               外呼下面有最小目标数3 => "中间变量2"."1号梯外呼下面有目标最小数3",
               外呼下面有最小目标数4 => "中间变量2"."1号梯外呼下面有目标最小数4",
               外呼下面有最小目标数5 => "中间变量2"."1号梯外呼下面有目标最小数5",
               外呼下面有最小目标数6 => "中间变量2"."1号梯外呼下面有目标最小数6",
               外呼下面有最小目标数7 => "中间变量2"."1号梯外呼下面有目标最小数7",
               外呼下面有最小目标数8 => "中间变量2"."1号梯外呼下面有目标最小数8",
               外呼下面有最小目标数9 => "中间变量2"."1号梯外呼下面有目标最小数9",
               外呼下面有最小目标数10 => "中间变量2"."1号梯外呼下面有目标最小数10");
   "2号梯有无目标判断"("1层上呼分配" := "中间变量2"."1层上呼分配2",   // "目标判断"
               "2层上呼分配" := "中间变量2"."2层上呼分配2",
               "2层下呼分配" := "中间变量2"."2层下呼分配2",
               "3层上呼分配" := "中间变量2"."3层上呼分配2",
               "3层下呼分配" := "中间变量2"."3层下呼分配2",
               "4层上呼分配" := "中间变量2"."4层上呼分配2",
               "4层下呼分配" := "中间变量2"."4层下呼分配2",
               "5层上呼分配" := "中间变量2"."5层上呼分配2",
               "5层下呼分配" := "中间变量2"."5层下呼分配2",
               "6层上呼分配" := "中间变量2"."6层上呼分配2",
               "6层下呼分配" := "中间变量2"."6层下呼分配2",
               "7层上呼分配" := "中间变量2"."7层上呼分配2",
               "7层下呼分配" := "中间变量2"."7层下呼分配2",
               "8层上呼分配" := "中间变量2"."8层上呼分配2",
               "8层下呼分配" := "中间变量2"."8层下呼分配2",
               "9层上呼分配" := "中间变量2"."9层上呼分配2",
               "9层下呼分配" := "中间变量2"."9层下呼分配2",
               "10层下呼分配" := "中间变量2"."10层下呼分配2",
               内呼按钮1 := "输出"."2号梯1层按钮指示灯",
               内呼按钮2 := "输出"."2号梯2层按钮指示灯",
               内呼按钮3 := "输出"."2号梯3层按钮指示灯",
               内呼按钮4 := "输出"."2号梯4层按钮指示灯",
               内呼按钮5 := "输出"."2号梯5层按钮指示灯",
               内呼按钮6 := "输出"."2号梯6层按钮指示灯",
               内呼按钮7 := "输出"."2号梯7层按钮指示灯",
               内呼按钮8 := "输出"."2号梯8层按钮指示灯",
               内呼按钮9 := "输出"."2号梯9层按钮指示灯",
               内呼按钮10 := "输出"."2号梯10层按钮指示灯",
               外呼下面无目标2 => "中间变量2"."2号梯外呼下面无目标2",
               外呼下面无目标3 => "中间变量2"."2号梯外呼下面无目标3",
               外呼下面无目标4 => "中间变量2"."2号梯外呼下面无目标4",
               外呼下面无目标5 => "中间变量2"."2号梯外呼下面无目标5",
               外呼下面无目标6 => "中间变量2"."2号梯外呼下面无目标6",
               外呼下面无目标7 => "中间变量2"."2号梯外呼下面无目标7",
               外呼下面无目标8 => "中间变量2"."2号梯外呼下面无目标8",
               外呼下面无目标9 => "中间变量2"."2号梯外呼下面无目标9",
               外呼上面无目标2 => "中间变量2"."2号梯外呼上面无目标2",
               外呼上面无目标3 => "中间变量2"."2号梯外呼上面无目标3",
               外呼上面无目标4 => "中间变量2"."2号梯外呼上面无目标4",
               外呼上面无目标5 => "中间变量2"."2号梯外呼上面无目标5",
               外呼上面无目标6 => "中间变量2"."2号梯外呼上面无目标6",
               外呼上面无目标7 => "中间变量2"."2号梯外呼上面无目标7",
               外呼上面无目标8 => "中间变量2"."2号梯外呼上面无目标8",
               外呼上面无目标9 => "中间变量2"."2号梯外呼上面无目标9",
               外呼上面有目标1 => "中间变量2"."2号梯外呼上面有目标1",
               外呼上面有目标2 => "中间变量2"."2号梯外呼上面有目标2",
               外呼上面有目标3 => "中间变量2"."2号梯外呼上面有目标3",
               外呼上面有目标4 => "中间变量2"."2号梯外呼上面有目标4",
               外呼上面有目标5 => "中间变量2"."2号梯外呼上面有目标5",
               外呼上面有目标6 => "中间变量2"."2号梯外呼上面有目标6",
               外呼上面有目标7 => "中间变量2"."2号梯外呼上面有目标7",
               外呼上面有目标8 => "中间变量2"."2号梯外呼上面有目标8",
               外呼上面有目标9 => "中间变量2"."2号梯外呼上面有目标9",
               外呼下面有目标2 => "中间变量2"."2号梯外呼下面有目标2",
               外呼下面有目标3 => "中间变量2"."2号梯外呼下面有目标3",
               外呼下面有目标4 => "中间变量2"."2号梯外呼下面有目标4",
               外呼下面有目标5 => "中间变量2"."2号梯外呼下面有目标5",
               外呼下面有目标6 => "中间变量2"."2号梯外呼下面有目标6",
               外呼下面有目标7 => "中间变量2"."2号梯外呼下面有目标7",
               外呼下面有目标8 => "中间变量2"."2号梯外呼下面有目标8",
               外呼下面有目标9 => "中间变量2"."2号梯外呼下面有目标9",
               外呼下面有目标10 => "中间变量2"."2号梯外呼下面有目标10",
               外呼上面有最大目标数1 => "中间变量2"."2号梯外呼上面有目标最大数1",
               外呼上面有最大目标数2 => "中间变量2"."2号梯外呼上面有目标最大数2",
               外呼上面有最大目标数3 => "中间变量2"."2号梯外呼上面有目标最大数3",
               外呼上面有最大目标数4 => "中间变量2"."2号梯外呼上面有目标最大数4",
               外呼上面有最大目标数5 => "中间变量2"."2号梯外呼上面有目标最大数5",
               外呼上面有最大目标数6 => "中间变量2"."2号梯外呼上面有目标最大数6",
               外呼上面有最大目标数7 => "中间变量2"."2号梯外呼上面有目标最大数7",
               外呼上面有最大目标数8 => "中间变量2"."2号梯外呼上面有目标最大数8",
               外呼上面有最大目标数9 => "中间变量2"."2号梯外呼上面有目标最大数9",
               外呼下面有最小目标数2 => "中间变量2"."2号梯外呼下面有目标最小数2",
               外呼下面有最小目标数3 => "中间变量2"."2号梯外呼下面有目标最小数3",
               外呼下面有最小目标数4 => "中间变量2"."2号梯外呼下面有目标最小数4",
               外呼下面有最小目标数5 => "中间变量2"."2号梯外呼下面有目标最小数5",
               外呼下面有最小目标数6 => "中间变量2"."2号梯外呼下面有目标最小数6",
               外呼下面有最小目标数7 => "中间变量2"."2号梯外呼下面有目标最小数7",
               外呼下面有最小目标数8 => "中间变量2"."2号梯外呼下面有目标最小数8",
               外呼下面有最小目标数9 => "中间变量2"."2号梯外呼下面有目标最小数9",
               外呼下面有最小目标数10 => "中间变量2"."2号梯外呼下面有目标最小数10");
   "3号梯有无目标判断"("1层上呼分配" := "中间变量2"."1层上呼分配3",   // "目标判断"
               "2层上呼分配" := "中间变量2"."2层上呼分配3",
               "2层下呼分配" := "中间变量2"."2层下呼分配3",
               "3层上呼分配" := "中间变量2"."3层上呼分配3",
               "3层下呼分配" := "中间变量2"."3层下呼分配3",
               "4层上呼分配" := "中间变量2"."4层上呼分配3",
               "4层下呼分配" := "中间变量2"."4层下呼分配3",
               "5层上呼分配" := "中间变量2"."5层上呼分配3",
               "5层下呼分配" := "中间变量2"."5层下呼分配3",
               "6层上呼分配" := "中间变量2"."6层上呼分配3",
               "6层下呼分配" := "中间变量2"."6层下呼分配3",
               "7层上呼分配" := "中间变量2"."7层上呼分配3",
               "7层下呼分配" := "中间变量2"."7层下呼分配3",
               "8层上呼分配" := "中间变量2"."8层上呼分配3",
               "8层下呼分配" := "中间变量2"."8层下呼分配3",
               "9层上呼分配" := "中间变量2"."9层上呼分配3",
               "9层下呼分配" := "中间变量2"."9层下呼分配3",
               "10层下呼分配" := "中间变量2"."10层下呼分配3",
               内呼按钮1 := "输出"."3号梯1层按钮指示灯",
               内呼按钮2 := "输出"."3号梯2层按钮指示灯",
               内呼按钮3 := "输出"."3号梯3层按钮指示灯",
               内呼按钮4 := "输出"."3号梯4层按钮指示灯",
               内呼按钮5 := "输出"."3号梯5层按钮指示灯",
               内呼按钮6 := "输出"."3号梯6层按钮指示灯",
               内呼按钮7 := "输出"."3号梯7层按钮指示灯",
               内呼按钮8 := "输出"."3号梯8层按钮指示灯",
               内呼按钮9 := "输出"."3号梯9层按钮指示灯",
               内呼按钮10 := "输出"."3号梯10层按钮指示灯",
               外呼下面无目标2 => "中间变量2"."3号梯外呼下面无目标2",
               外呼下面无目标3 => "中间变量2"."3号梯外呼下面无目标3",
               外呼下面无目标4 => "中间变量2"."3号梯外呼下面无目标4",
               外呼下面无目标5 => "中间变量2"."3号梯外呼下面无目标5",
               外呼下面无目标6 => "中间变量2"."3号梯外呼下面无目标6",
               外呼下面无目标7 => "中间变量2"."3号梯外呼下面无目标7",
               外呼下面无目标8 => "中间变量2"."3号梯外呼下面无目标8",
               外呼下面无目标9 => "中间变量2"."3号梯外呼下面无目标9",
               外呼上面无目标2 => "中间变量2"."3号梯外呼上面无目标2",
               外呼上面无目标3 => "中间变量2"."3号梯外呼上面无目标3",
               外呼上面无目标4 => "中间变量2"."3号梯外呼上面无目标4",
               外呼上面无目标5 => "中间变量2"."3号梯外呼上面无目标5",
               外呼上面无目标6 => "中间变量2"."3号梯外呼上面无目标6",
               外呼上面无目标7 => "中间变量2"."3号梯外呼上面无目标7",
               外呼上面无目标8 => "中间变量2"."3号梯外呼上面无目标8",
               外呼上面无目标9 => "中间变量2"."3号梯外呼上面无目标9",
               外呼上面有目标1 => "中间变量2"."3号梯外呼上面有目标1",
               外呼上面有目标2 => "中间变量2"."3号梯外呼上面有目标2",
               外呼上面有目标3 => "中间变量2"."3号梯外呼上面有目标3",
               外呼上面有目标4 => "中间变量2"."3号梯外呼上面有目标4",
               外呼上面有目标5 => "中间变量2"."3号梯外呼上面有目标5",
               外呼上面有目标6 => "中间变量2"."3号梯外呼上面有目标6",
               外呼上面有目标7 => "中间变量2"."3号梯外呼上面有目标7",
               外呼上面有目标8 => "中间变量2"."3号梯外呼上面有目标8",
               外呼上面有目标9 => "中间变量2"."3号梯外呼上面有目标9",
               外呼下面有目标2 => "中间变量2"."3号梯外呼下面有目标2",
               外呼下面有目标3 => "中间变量2"."3号梯外呼下面有目标3",
               外呼下面有目标4 => "中间变量2"."3号梯外呼下面有目标4",
               外呼下面有目标5 => "中间变量2"."3号梯外呼下面有目标5",
               外呼下面有目标6 => "中间变量2"."3号梯外呼下面有目标6",
               外呼下面有目标7 => "中间变量2"."3号梯外呼下面有目标7",
               外呼下面有目标8 => "中间变量2"."3号梯外呼下面有目标8",
               外呼下面有目标9 => "中间变量2"."3号梯外呼下面有目标9",
               外呼下面有目标10 => "中间变量2"."3号梯外呼下面有目标10",
               外呼上面有最大目标数1 => "中间变量2"."3号梯外呼上面有目标最大数1",
               外呼上面有最大目标数2 => "中间变量2"."3号梯外呼上面有目标最大数2",
               外呼上面有最大目标数3 => "中间变量2"."3号梯外呼上面有目标最大数3",
               外呼上面有最大目标数4 => "中间变量2"."3号梯外呼上面有目标最大数4",
               外呼上面有最大目标数5 => "中间变量2"."3号梯外呼上面有目标最大数5",
               外呼上面有最大目标数6 => "中间变量2"."3号梯外呼上面有目标最大数6",
               外呼上面有最大目标数7 => "中间变量2"."3号梯外呼上面有目标最大数7",
               外呼上面有最大目标数8 => "中间变量2"."3号梯外呼上面有目标最大数8",
               外呼上面有最大目标数9 => "中间变量2"."3号梯外呼上面有目标最大数9",
               外呼下面有最小目标数2 => "中间变量2"."3号梯外呼下面有目标最小数2",
               外呼下面有最小目标数3 => "中间变量2"."3号梯外呼下面有目标最小数3",
               外呼下面有最小目标数4 => "中间变量2"."3号梯外呼下面有目标最小数4",
               外呼下面有最小目标数5 => "中间变量2"."3号梯外呼下面有目标最小数5",
               外呼下面有最小目标数6 => "中间变量2"."3号梯外呼下面有目标最小数6",
               外呼下面有最小目标数7 => "中间变量2"."3号梯外呼下面有目标最小数7",
               外呼下面有最小目标数8 => "中间变量2"."3号梯外呼下面有目标最小数8",
               外呼下面有最小目标数9 => "中间变量2"."3号梯外呼下面有目标最小数9",
               外呼下面有最小目标数10 => "中间变量2"."3号梯外呼下面有目标最小数10");
   "4号梯有无目标判断"("1层上呼分配" := "中间变量2"."1层上呼分配4",   // "目标判断"
               "2层上呼分配" := "中间变量2"."2层上呼分配4",
               "2层下呼分配" := "中间变量2"."2层下呼分配4",
               "3层上呼分配" := "中间变量2"."3层上呼分配4",
               "3层下呼分配" := "中间变量2"."3层下呼分配4",
               "4层上呼分配" := "中间变量2"."4层上呼分配4",
               "4层下呼分配" := "中间变量2"."4层下呼分配4",
               "5层上呼分配" := "中间变量2"."5层上呼分配4",
               "5层下呼分配" := "中间变量2"."5层下呼分配4",
               "6层上呼分配" := "中间变量2"."6层上呼分配4",
               "6层下呼分配" := "中间变量2"."6层下呼分配4",
               "7层上呼分配" := "中间变量2"."7层上呼分配4",
               "7层下呼分配" := "中间变量2"."7层下呼分配4",
               "8层上呼分配" := "中间变量2"."8层上呼分配4",
               "8层下呼分配" := "中间变量2"."8层下呼分配4",
               "9层上呼分配" := "中间变量2"."9层上呼分配4",
               "9层下呼分配" := "中间变量2"."9层下呼分配4",
               "10层下呼分配" := "中间变量2"."10层下呼分配4",
               内呼按钮1 := "输出"."4号梯1层按钮指示灯",
               内呼按钮2 := "输出"."4号梯2层按钮指示灯",
               内呼按钮3 := "输出"."4号梯3层按钮指示灯",
               内呼按钮4 := "输出"."4号梯4层按钮指示灯",
               内呼按钮5 := "输出"."4号梯5层按钮指示灯",
               内呼按钮6 := "输出"."4号梯6层按钮指示灯",
               内呼按钮7 := "输出"."4号梯7层按钮指示灯",
               内呼按钮8 := "输出"."4号梯8层按钮指示灯",
               内呼按钮9 := "输出"."4号梯9层按钮指示灯",
               内呼按钮10 := "输出"."4号梯10层按钮指示灯",
               外呼下面无目标2 => "中间变量2"."4号梯外呼下面无目标2",
               外呼下面无目标3 => "中间变量2"."4号梯外呼下面无目标3",
               外呼下面无目标4 => "中间变量2"."4号梯外呼下面无目标4",
               外呼下面无目标5 => "中间变量2"."4号梯外呼下面无目标5",
               外呼下面无目标6 => "中间变量2"."4号梯外呼下面无目标6",
               外呼下面无目标7 => "中间变量2"."4号梯外呼下面无目标7",
               外呼下面无目标8 => "中间变量2"."4号梯外呼下面无目标8",
               外呼下面无目标9 => "中间变量2"."4号梯外呼下面无目标9",
               外呼上面无目标2 => "中间变量2"."4号梯外呼上面无目标2",
               外呼上面无目标3 => "中间变量2"."4号梯外呼上面无目标3",
               外呼上面无目标4 => "中间变量2"."4号梯外呼上面无目标4",
               外呼上面无目标5 => "中间变量2"."4号梯外呼上面无目标5",
               外呼上面无目标6 => "中间变量2"."4号梯外呼上面无目标6",
               外呼上面无目标7 => "中间变量2"."4号梯外呼上面无目标7",
               外呼上面无目标8 => "中间变量2"."4号梯外呼上面无目标8",
               外呼上面无目标9 => "中间变量2"."4号梯外呼上面无目标9",
               外呼上面有目标1 => "中间变量2"."4号梯外呼上面有目标1",
               外呼上面有目标2 => "中间变量2"."4号梯外呼上面有目标2",
               外呼上面有目标3 => "中间变量2"."4号梯外呼上面有目标3",
               外呼上面有目标4 => "中间变量2"."4号梯外呼上面有目标4",
               外呼上面有目标5 => "中间变量2"."4号梯外呼上面有目标5",
               外呼上面有目标6 => "中间变量2"."4号梯外呼上面有目标6",
               外呼上面有目标7 => "中间变量2"."4号梯外呼上面有目标7",
               外呼上面有目标8 => "中间变量2"."4号梯外呼上面有目标8",
               外呼上面有目标9 => "中间变量2"."4号梯外呼上面有目标9",
               外呼下面有目标2 => "中间变量2"."4号梯外呼下面有目标2",
               外呼下面有目标3 => "中间变量2"."4号梯外呼下面有目标3",
               外呼下面有目标4 => "中间变量2"."4号梯外呼下面有目标4",
               外呼下面有目标5 => "中间变量2"."4号梯外呼下面有目标5",
               外呼下面有目标6 => "中间变量2"."4号梯外呼下面有目标6",
               外呼下面有目标7 => "中间变量2"."4号梯外呼下面有目标7",
               外呼下面有目标8 => "中间变量2"."4号梯外呼下面有目标8",
               外呼下面有目标9 => "中间变量2"."4号梯外呼下面有目标9",
               外呼下面有目标10 => "中间变量2"."4号梯外呼下面有目标10",
               外呼上面有最大目标数1 => "中间变量2"."4号梯外呼上面有目标最大数1",
               外呼上面有最大目标数2 => "中间变量2"."4号梯外呼上面有目标最大数2",
               外呼上面有最大目标数3 => "中间变量2"."4号梯外呼上面有目标最大数3",
               外呼上面有最大目标数4 => "中间变量2"."4号梯外呼上面有目标最大数4",
               外呼上面有最大目标数5 => "中间变量2"."4号梯外呼上面有目标最大数5",
               外呼上面有最大目标数6 => "中间变量2"."4号梯外呼上面有目标最大数6",
               外呼上面有最大目标数7 => "中间变量2"."4号梯外呼上面有目标最大数7",
               外呼上面有最大目标数8 => "中间变量2"."4号梯外呼上面有目标最大数8",
               外呼上面有最大目标数9 => "中间变量2"."4号梯外呼上面有目标最大数9",
               外呼下面有最小目标数2 => "中间变量2"."4号梯外呼下面有目标最小数2",
               外呼下面有最小目标数3 => "中间变量2"."4号梯外呼下面有目标最小数3",
               外呼下面有最小目标数4 => "中间变量2"."4号梯外呼下面有目标最小数4",
               外呼下面有最小目标数5 => "中间变量2"."4号梯外呼下面有目标最小数5",
               外呼下面有最小目标数6 => "中间变量2"."4号梯外呼下面有目标最小数6",
               外呼下面有最小目标数7 => "中间变量2"."4号梯外呼下面有目标最小数7",
               外呼下面有最小目标数8 => "中间变量2"."4号梯外呼下面有目标最小数8",
               外呼下面有最小目标数9 => "中间变量2"."4号梯外呼下面有目标最小数9",
               外呼下面有最小目标数10 => "中间变量2"."4号梯外呼下面有目标最小数10");
   "5号梯有无目标判断"("1层上呼分配" := "中间变量2"."1层上呼分配5",   // "目标判断"
               "2层上呼分配" := "中间变量2"."2层上呼分配5",
               "2层下呼分配" := "中间变量2"."2层下呼分配5",
               "3层上呼分配" := "中间变量2"."3层上呼分配5",
               "3层下呼分配" := "中间变量2"."3层下呼分配5",
               "4层上呼分配" := "中间变量2"."4层上呼分配5",
               "4层下呼分配" := "中间变量2"."4层下呼分配5",
               "5层上呼分配" := "中间变量2"."5层上呼分配5",
               "5层下呼分配" := "中间变量2"."5层下呼分配5",
               "6层上呼分配" := "中间变量2"."6层上呼分配5",
               "6层下呼分配" := "中间变量2"."6层下呼分配5",
               "7层上呼分配" := "中间变量2"."7层上呼分配5",
               "7层下呼分配" := "中间变量2"."7层下呼分配5",
               "8层上呼分配" := "中间变量2"."8层上呼分配5",
               "8层下呼分配" := "中间变量2"."8层下呼分配5",
               "9层上呼分配" := "中间变量2"."9层上呼分配5",
               "9层下呼分配" := "中间变量2"."9层下呼分配5",
               "10层下呼分配" := "中间变量2"."10层下呼分配5",
               内呼按钮1 := "输出"."5号梯1层按钮指示灯",
               内呼按钮2 := "输出"."5号梯2层按钮指示灯",
               内呼按钮3 := "输出"."5号梯3层按钮指示灯",
               内呼按钮4 := "输出"."5号梯4层按钮指示灯",
               内呼按钮5 := "输出"."5号梯5层按钮指示灯",
               内呼按钮6 := "输出"."5号梯6层按钮指示灯",
               内呼按钮7 := "输出"."5号梯7层按钮指示灯",
               内呼按钮8 := "输出"."5号梯8层按钮指示灯",
               内呼按钮9 := "输出"."5号梯9层按钮指示灯",
               内呼按钮10 := "输出"."5号梯10层按钮指示灯",
               外呼下面无目标2 => "中间变量2"."5号梯外呼下面无目标2",
               外呼下面无目标3 => "中间变量2"."5号梯外呼下面无目标3",
               外呼下面无目标4 => "中间变量2"."5号梯外呼下面无目标4",
               外呼下面无目标5 => "中间变量2"."5号梯外呼下面无目标5",
               外呼下面无目标6 => "中间变量2"."5号梯外呼下面无目标6",
               外呼下面无目标7 => "中间变量2"."5号梯外呼下面无目标7",
               外呼下面无目标8 => "中间变量2"."5号梯外呼下面无目标8",
               外呼下面无目标9 => "中间变量2"."5号梯外呼下面无目标9",
               外呼上面无目标2 => "中间变量2"."5号梯外呼上面无目标2",
               外呼上面无目标3 => "中间变量2"."5号梯外呼上面无目标3",
               外呼上面无目标4 => "中间变量2"."5号梯外呼上面无目标4",
               外呼上面无目标5 => "中间变量2"."5号梯外呼上面无目标5",
               外呼上面无目标6 => "中间变量2"."5号梯外呼上面无目标6",
               外呼上面无目标7 => "中间变量2"."5号梯外呼上面无目标7",
               外呼上面无目标8 => "中间变量2"."5号梯外呼上面无目标8",
               外呼上面无目标9 => "中间变量2"."5号梯外呼上面无目标9",
               外呼上面有目标1 => "中间变量2"."5号梯外呼上面有目标1",
               外呼上面有目标2 => "中间变量2"."5号梯外呼上面有目标2",
               外呼上面有目标3 => "中间变量2"."5号梯外呼上面有目标3",
               外呼上面有目标4 => "中间变量2"."5号梯外呼上面有目标4",
               外呼上面有目标5 => "中间变量2"."5号梯外呼上面有目标5",
               外呼上面有目标6 => "中间变量2"."5号梯外呼上面有目标6",
               外呼上面有目标7 => "中间变量2"."5号梯外呼上面有目标7",
               外呼上面有目标8 => "中间变量2"."5号梯外呼上面有目标8",
               外呼上面有目标9 => "中间变量2"."5号梯外呼上面有目标9",
               外呼下面有目标2 => "中间变量2"."5号梯外呼下面有目标2",
               外呼下面有目标3 => "中间变量2"."5号梯外呼下面有目标3",
               外呼下面有目标4 => "中间变量2"."5号梯外呼下面有目标4",
               外呼下面有目标5 => "中间变量2"."5号梯外呼下面有目标5",
               外呼下面有目标6 => "中间变量2"."5号梯外呼下面有目标6",
               外呼下面有目标7 => "中间变量2"."5号梯外呼下面有目标7",
               外呼下面有目标8 => "中间变量2"."5号梯外呼下面有目标8",
               外呼下面有目标9 => "中间变量2"."5号梯外呼下面有目标9",
               外呼下面有目标10 => "中间变量2"."5号梯外呼下面有目标10",
               外呼上面有最大目标数1 => "中间变量2"."5号梯外呼上面有目标最大数1",
               外呼上面有最大目标数2 => "中间变量2"."5号梯外呼上面有目标最大数2",
               外呼上面有最大目标数3 => "中间变量2"."5号梯外呼上面有目标最大数3",
               外呼上面有最大目标数4 => "中间变量2"."5号梯外呼上面有目标最大数4",
               外呼上面有最大目标数5 => "中间变量2"."5号梯外呼上面有目标最大数5",
               外呼上面有最大目标数6 => "中间变量2"."5号梯外呼上面有目标最大数6",
               外呼上面有最大目标数7 => "中间变量2"."5号梯外呼上面有目标最大数7",
               外呼上面有最大目标数8 => "中间变量2"."5号梯外呼上面有目标最大数8",
               外呼上面有最大目标数9 => "中间变量2"."5号梯外呼上面有目标最大数9",
               外呼下面有最小目标数2 => "中间变量2"."5号梯外呼下面有目标最小数2",
               外呼下面有最小目标数3 => "中间变量2"."5号梯外呼下面有目标最小数3",
               外呼下面有最小目标数4 => "中间变量2"."5号梯外呼下面有目标最小数4",
               外呼下面有最小目标数5 => "中间变量2"."5号梯外呼下面有目标最小数5",
               外呼下面有最小目标数6 => "中间变量2"."5号梯外呼下面有目标最小数6",
               外呼下面有最小目标数7 => "中间变量2"."5号梯外呼下面有目标最小数7",
               外呼下面有最小目标数8 => "中间变量2"."5号梯外呼下面有目标最小数8",
               外呼下面有最小目标数9 => "中间变量2"."5号梯外呼下面有目标最小数9",
               外呼下面有最小目标数10 => "中间变量2"."5号梯外呼下面有目标最小数10");
   "6号梯有无目标判断"("1层上呼分配" := "中间变量2"."1层上呼分配6",   // "目标判断"
               "2层上呼分配" := "中间变量2"."2层上呼分配6",
               "2层下呼分配" := "中间变量2"."2层下呼分配6",
               "3层上呼分配" := "中间变量2"."3层上呼分配6",
               "3层下呼分配" := "中间变量2"."3层下呼分配6",
               "4层上呼分配" := "中间变量2"."4层上呼分配6",
               "4层下呼分配" := "中间变量2"."4层下呼分配6",
               "5层上呼分配" := "中间变量2"."5层上呼分配6",
               "5层下呼分配" := "中间变量2"."5层下呼分配6",
               "6层上呼分配" := "中间变量2"."6层上呼分配6",
               "6层下呼分配" := "中间变量2"."6层下呼分配6",
               "7层上呼分配" := "中间变量2"."7层上呼分配6",
               "7层下呼分配" := "中间变量2"."7层下呼分配6",
               "8层上呼分配" := "中间变量2"."8层上呼分配6",
               "8层下呼分配" := "中间变量2"."8层下呼分配6",
               "9层上呼分配" := "中间变量2"."9层上呼分配6",
               "9层下呼分配" := "中间变量2"."9层下呼分配6",
               "10层下呼分配" := "中间变量2"."10层下呼分配6",
               内呼按钮1 := "输出"."6号梯1层按钮指示灯",
               内呼按钮2 := "输出"."6号梯2层按钮指示灯",
               内呼按钮3 := "输出"."6号梯3层按钮指示灯",
               内呼按钮4 := "输出"."6号梯4层按钮指示灯",
               内呼按钮5 := "输出"."6号梯5层按钮指示灯",
               内呼按钮6 := "输出"."6号梯6层按钮指示灯",
               内呼按钮7 := "输出"."6号梯7层按钮指示灯",
               内呼按钮8 := "输出"."6号梯8层按钮指示灯",
               内呼按钮9 := "输出"."6号梯9层按钮指示灯",
               内呼按钮10 := "输出"."6号梯10层按钮指示灯",
               外呼下面无目标2 => "中间变量2"."6号梯外呼下面无目标2",
               外呼下面无目标3 => "中间变量2"."6号梯外呼下面无目标3",
               外呼下面无目标4 => "中间变量2"."6号梯外呼下面无目标4",
               外呼下面无目标5 => "中间变量2"."6号梯外呼下面无目标5",
               外呼下面无目标6 => "中间变量2"."6号梯外呼下面无目标6",
               外呼下面无目标7 => "中间变量2"."6号梯外呼下面无目标7",
               外呼下面无目标8 => "中间变量2"."6号梯外呼下面无目标8",
               外呼下面无目标9 => "中间变量2"."6号梯外呼下面无目标9",
               外呼上面无目标2 => "中间变量2"."6号梯外呼上面无目标2",
               外呼上面无目标3 => "中间变量2"."6号梯外呼上面无目标3",
               外呼上面无目标4 => "中间变量2"."6号梯外呼上面无目标4",
               外呼上面无目标5 => "中间变量2"."6号梯外呼上面无目标5",
               外呼上面无目标6 => "中间变量2"."6号梯外呼上面无目标6",
               外呼上面无目标7 => "中间变量2"."6号梯外呼上面无目标7",
               外呼上面无目标8 => "中间变量2"."6号梯外呼上面无目标8",
               外呼上面无目标9 => "中间变量2"."6号梯外呼上面无目标9",
               外呼上面有目标1 => "中间变量2"."6号梯外呼上面有目标1",
               外呼上面有目标2 => "中间变量2"."6号梯外呼上面有目标2",
               外呼上面有目标3 => "中间变量2"."6号梯外呼上面有目标3",
               外呼上面有目标4 => "中间变量2"."6号梯外呼上面有目标4",
               外呼上面有目标5 => "中间变量2"."6号梯外呼上面有目标5",
               外呼上面有目标6 => "中间变量2"."6号梯外呼上面有目标6",
               外呼上面有目标7 => "中间变量2"."6号梯外呼上面有目标7",
               外呼上面有目标8 => "中间变量2"."6号梯外呼上面有目标8",
               外呼上面有目标9 => "中间变量2"."6号梯外呼上面有目标9",
               外呼下面有目标2 => "中间变量2"."6号梯外呼下面有目标2",
               外呼下面有目标3 => "中间变量2"."6号梯外呼下面有目标3",
               外呼下面有目标4 => "中间变量2"."6号梯外呼下面有目标4",
               外呼下面有目标5 => "中间变量2"."6号梯外呼下面有目标5",
               外呼下面有目标6 => "中间变量2"."6号梯外呼下面有目标6",
               外呼下面有目标7 => "中间变量2"."6号梯外呼下面有目标7",
               外呼下面有目标8 => "中间变量2"."6号梯外呼下面有目标8",
               外呼下面有目标9 => "中间变量2"."6号梯外呼下面有目标9",
               外呼下面有目标10 => "中间变量2"."6号梯外呼下面有目标10",
               外呼上面有最大目标数1 => "中间变量2"."6号梯外呼上面有目标最大数1",
               外呼上面有最大目标数2 => "中间变量2"."6号梯外呼上面有目标最大数2",
               外呼上面有最大目标数3 => "中间变量2"."6号梯外呼上面有目标最大数3",
               外呼上面有最大目标数4 => "中间变量2"."6号梯外呼上面有目标最大数4",
               外呼上面有最大目标数5 => "中间变量2"."6号梯外呼上面有目标最大数5",
               外呼上面有最大目标数6 => "中间变量2"."6号梯外呼上面有目标最大数6",
               外呼上面有最大目标数7 => "中间变量2"."6号梯外呼上面有目标最大数7",
               外呼上面有最大目标数8 => "中间变量2"."6号梯外呼上面有目标最大数8",
               外呼上面有最大目标数9 => "中间变量2"."6号梯外呼上面有目标最大数9",
               外呼下面有最小目标数2 => "中间变量2"."6号梯外呼下面有目标最小数2",
               外呼下面有最小目标数3 => "中间变量2"."6号梯外呼下面有目标最小数3",
               外呼下面有最小目标数4 => "中间变量2"."6号梯外呼下面有目标最小数4",
               外呼下面有最小目标数5 => "中间变量2"."6号梯外呼下面有目标最小数5",
               外呼下面有最小目标数6 => "中间变量2"."6号梯外呼下面有目标最小数6",
               外呼下面有最小目标数7 => "中间变量2"."6号梯外呼下面有目标最小数7",
               外呼下面有最小目标数8 => "中间变量2"."6号梯外呼下面有目标最小数8",
               外呼下面有最小目标数9 => "中间变量2"."6号梯外呼下面有目标最小数9",
               外呼下面有最小目标数10 => "中间变量2"."6号梯外呼下面有目标最小数10");
END_REGION
END_FUNCTION

FUNCTION "***********" : Void   // FC13, SCL
{ S7_Optimized_Access := 'TRUE' }
VERSION : 0.1
BEGIN
   //------------------------------------------------------------------
   //电梯运行中故障是否在最近楼层开门，还是直接停止运行？
   //1，最近楼层开门：外呼分配复位，突然检修信号置位，低速接触器置位，高速接触器复位，待上下平层=1后，电机，上下行接触器，高低速接触器复位，开门信号保持
   //2，直接停止运行：外呼分配复位，电机启动信号复位，上下行接触器复位，高低速接触器复位
   //------------------------------------------------------------------
   //减速控制，一级制动，二级制动，三级制动设置？
   //在电梯到达目标层前一层提供准备刹车信号，在电梯上行时，当上平层信号为1，电梯进行一级制动，在上下平层同时置位时，进行2级制动，100ms后进行三级制动。
   //------------------------------------------------------------------
   //开门超过一定时间后能否强行关门？
   //不可行，因为万一满载信号有，但电梯不能启动，就卡死
   //------------------------------------------------------------------
   //初始化检修完成后，在运行过程中检修复位，运行方向？
   //也在初始化赋值里调
   //------------------------------------------------------------------
   //在1层时下行接触器复位，在10层时上行接触器复位是否完成？
   //完成
   //------------------------------------------------------------------
   //开始后先修改：1、最大载重量 2、电梯初始化运行方向 3、初始化楼层数 4、初始化速度
   //------------------------------------------------------------------
   //在初始化时，上下行指示灯亮，数码管不亮
   //在初始化可以将上下行指示连到上下行指示灯上，在初始化完成后复位。
   //------------------------------------------------------------------
   //超重后故障指示灯是否亮？
   //
   //------------------------------------------------------------------
   //初始化时间过长/上下行指示灯闪烁？？
   //------------------------------------------------------------------
   //wincc 电梯状态画面按钮为绿色（已改）
END_FUNCTION

FUNCTION "程序运行时长" : Void   // FC14, LAD
{ S7_Optimized_Access := 'TRUE' }
VERSION : 0.1
   VAR_TEMP
      tag : Time;
      置位触发器 : Bool;
      tag1 : Bool;
      tag2 : Bool;
   END_VAR
   VAR CONSTANT
      开始信号 : Bool := 1;
   END_VAR
   VAR_TEMP   // added for the SCL form of the ladder/FBD networks
      _w1 : Bool;
      _w2 : Bool;
   END_VAR
BEGIN

REGION Network 1
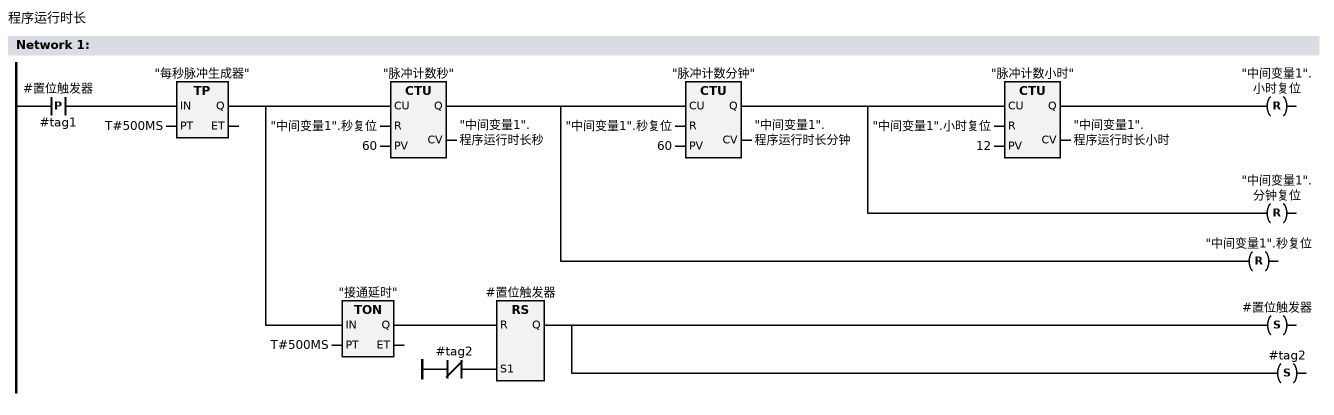
   #_w1 := #置位触发器 AND NOT #tag1;   // rising edge of #置位触发器
   #tag1 := #置位触发器;
   "每秒脉冲生成器".TP(IN := #_w1, PT := T#500MS);
   "脉冲计数秒".CTU(CU := "每秒脉冲生成器".Q, R := "中间变量1".秒复位, PV := 60, CV => "中间变量1".程序运行时长秒);
   "脉冲计数分钟".CTU(CU := "脉冲计数秒".Q, R := "中间变量1".秒复位, PV := 60, CV => "中间变量1".程序运行时长分钟);
   "脉冲计数小时".CTU(CU := "脉冲计数分钟".Q, R := "中间变量1".小时复位, PV := 12, CV => "中间变量1".程序运行时长小时);
   IF "脉冲计数小时".Q THEN "中间变量1".小时复位 := FALSE; END_IF;
   IF "脉冲计数分钟".Q THEN "中间变量1".分钟复位 := FALSE; END_IF;
   IF "脉冲计数秒".Q THEN "中间变量1".秒复位 := FALSE; END_IF;
   "接通延时".TON(IN := "每秒脉冲生成器".Q, PT := T#500MS);
   IF "接通延时".Q THEN
       #置位触发器 := FALSE;   // RS flip-flop
   END_IF;
   IF NOT #tag2 THEN #置位触发器 := TRUE; END_IF;
   #_w2 := #置位触发器;
   IF #_w2 THEN
       #置位触发器 := TRUE;
       #tag2 := TRUE;
   END_IF;
END_REGION
END_FUNCTION

ORGANIZATION_BLOCK "Main"   // OB1, LAD, ProgramCycle
TITLE = "Main Program Sweep (Cycle)"
{ S7_Optimized_Access := 'TRUE' }
VERSION : 0.1
   VAR_INPUT
      Initial_Call : Bool;   // Initial call of this OB
      Remanence : Bool;   // =True, if remanent data are available
   END_VAR
BEGIN

REGION Network 1: 程序运行时长
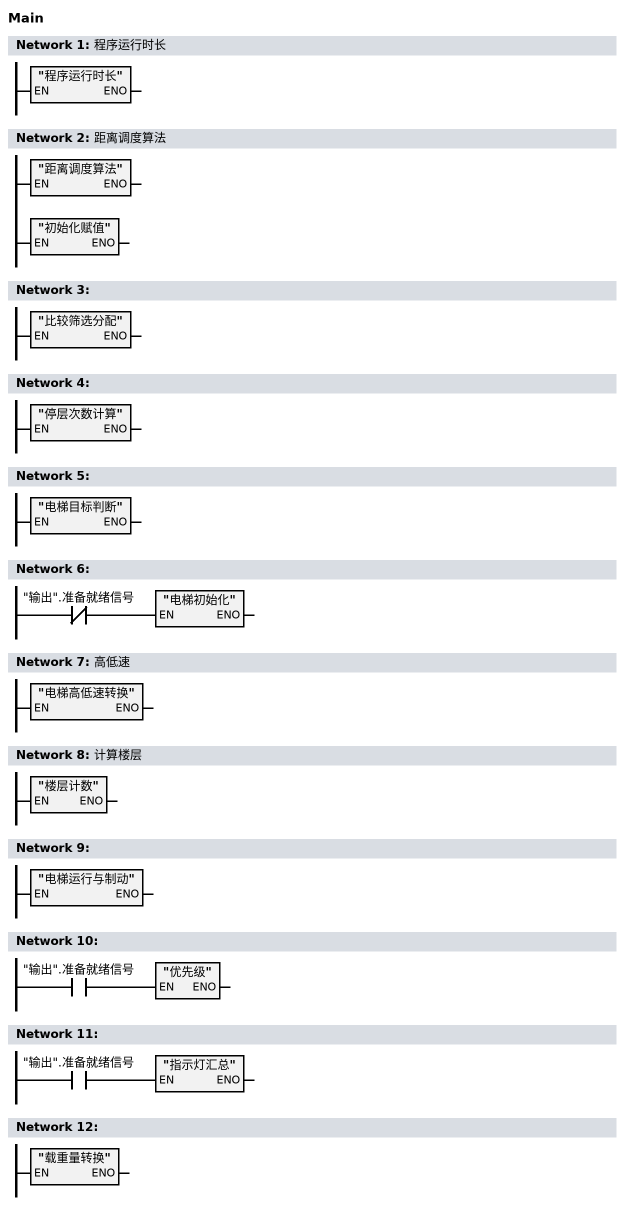
   RUNG wire#powerrail
      "程序运行时长"()
   END_RUNG
   // the same network as SCL:
   "程序运行时长"();
END_REGION

REGION Network 2: 距离调度算法
   RUNG wire#powerrail
      "距离调度算法"()
   END_RUNG
   RUNG wire#powerrail
      "初始化赋值"()
   END_RUNG
   // the same network as SCL:
   "距离调度算法"();
   "初始化赋值"();
END_REGION

REGION Network 3
   RUNG wire#powerrail
      "比较筛选分配"()
   END_RUNG
   // the same network as SCL:
   "比较筛选分配"();
END_REGION

REGION Network 4
   RUNG wire#powerrail
      "停层次数计算"()
   END_RUNG
   // the same network as SCL:
   "停层次数计算"();
END_REGION

REGION Network 5
   RUNG wire#powerrail
      "电梯目标判断"()
   END_RUNG
   // the same network as SCL:
   "电梯目标判断"();
END_REGION

REGION Network 6
   RUNG wire#powerrail
      I_Contact( "输出".准备就绪信号 )
      "电梯初始化"()
   END_RUNG
   // the same network as SCL:
   IF NOT "输出".准备就绪信号 THEN "电梯初始化"(); END_IF;
END_REGION

REGION Network 7: 高低速
   RUNG wire#powerrail
      "电梯高低速转换"()
   END_RUNG
   // the same network as SCL:
   "电梯高低速转换"();
END_REGION

REGION Network 8: 计算楼层
   RUNG wire#powerrail
      "楼层计数"()
   END_RUNG
   // the same network as SCL:
   "楼层计数"();
END_REGION

REGION Network 9
   RUNG wire#powerrail
      "电梯运行与制动"()
   END_RUNG
   // the same network as SCL:
   "电梯运行与制动"();
END_REGION

REGION Network 10
   RUNG wire#powerrail
      Contact( "输出".准备就绪信号 )
      "优先级"()
   END_RUNG
   // the same network as SCL:
   IF "输出".准备就绪信号 THEN "优先级"(); END_IF;
END_REGION

REGION Network 11
   RUNG wire#powerrail
      Contact( "输出".准备就绪信号 )
      "指示灯汇总"()
   END_RUNG
   // the same network as SCL:
   IF "输出".准备就绪信号 THEN "指示灯汇总"(); END_IF;
END_REGION

REGION Network 12
   RUNG wire#powerrail
      "载重量转换"()
   END_RUNG
   // the same network as SCL:
   "载重量转换"();
END_REGION
END_ORGANIZATION_BLOCK

(* ===== HMI "HMI_RT_1" =====
system functions are stored by id; their names below are inferred from use
connection "HMI__1": ETHERNET, S7_1200_OMS

HMI tags "默认变量表"
   "密码" : WString[254], internal
   "当前用户名" : WString[254], internal
   "提示信息" : WString[254], internal
   "用户名" : WString[254], internal
   "用户名或密码错误" : WString[254], internal
   "用户未登录" : WString[254], internal
   "登录成功" : WString[254], internal
   "当前运行时间" : WString[254], internal
      on ChangeValue: function_e3503463('record.csv', U 0, 2, 1, N)

HMI tags "默认变量表1"
   "输入_1层上行呼梯按钮" : Bool = PLC 输入.1层上行呼梯按钮 AT %DB10.DBX0.0, 100 ms
   "输入_2层上行呼梯按钮" : Bool = PLC 输入.2层上行呼梯按钮 AT %DB10.DBX0.1, 100 ms
   "输入_3层上行呼梯按钮" : Bool = PLC 输入.3层上行呼梯按钮 AT %DB10.DBX0.2, 100 ms
   "输入_4层上行呼梯按钮" : Bool = PLC 输入.4层上行呼梯按钮 AT %DB10.DBX0.3, 100 ms
   "输入_5层上行呼梯按钮" : Bool = PLC 输入.5层上行呼梯按钮 AT %DB10.DBX0.4, 100 ms
   "输入_6层上行呼梯按钮" : Bool = PLC 输入.6层上行呼梯按钮 AT %DB10.DBX0.5, 100 ms
   "输入_7层上行呼梯按钮" : Bool = PLC 输入.7层上行呼梯按钮 AT %DB10.DBX0.6, 100 ms
   "输入_8层上行呼梯按钮" : Bool = PLC 输入.8层上行呼梯按钮 AT %DB10.DBX0.7, 100 ms
   "输入_9层上行呼梯按钮" : Bool = PLC 输入.9层上行呼梯按钮 AT %DB10.DBX1.0, 100 ms
   "输入_10层下行呼梯按钮" : Bool = PLC 输入.10层下行呼梯按钮 AT %DB10.DBX2.1, 100 ms
   "输入_3层下行呼梯按钮" : Bool = PLC 输入.3层下行呼梯按钮 AT %DB10.DBX1.2, 100 ms
   "输入_4层下行呼梯按钮" : Bool = PLC 输入.4层下行呼梯按钮 AT %DB10.DBX1.3, 100 ms
   "输入_5层下行呼梯按钮" : Bool = PLC 输入.5层下行呼梯按钮 AT %DB10.DBX1.4, 100 ms
   "输入_6层下行呼梯按钮" : Bool = PLC 输入.6层下行呼梯按钮 AT %DB10.DBX1.5, 100 ms
   "输入_7层下行呼梯按钮" : Bool = PLC 输入.7层下行呼梯按钮 AT %DB10.DBX1.6, 100 ms
   "输入_8层下行呼梯按钮" : Bool = PLC 输入.8层下行呼梯按钮 AT %DB10.DBX1.7, 100 ms
   "输入_9层下行呼梯按钮" : Bool = PLC 输入.9层下行呼梯按钮 AT %DB10.DBX2.0, 100 ms
   "输入_自动运行信号" : Bool = PLC 输入.自动运行信号 AT %DB10.DBX27.0, 100 ms
   "输出_1号梯满载指示" : Bool = PLC 输出.1号梯满载指示 AT %DB11.DBX5.7, 100 ms
   "输出_1号梯故障指示" : Bool = PLC 输出.1号梯故障指示 AT %DB11.DBX5.4, 100 ms
   "输出_准备就绪信号" : Bool = PLC 输出.准备就绪信号 AT %DB11.DBX32.2, 100 ms
   "输出_1号梯照明指示" : Bool = PLC 输出.1号梯照明指示 AT %DB11.DBX5.5, 100 ms
   "输出_1号梯风扇指示" : Bool = PLC 输出.1号梯风扇指示 AT %DB11.DBX5.6, 100 ms
   "输入_1号梯轿内选层按钮1" : Bool = PLC 输入.1号梯轿内选层按钮1 AT %DB10.DBX2.2, 100 ms
   "输入_1号梯轿内选层按钮2" : Bool = PLC 输入.1号梯轿内选层按钮2 AT %DB10.DBX2.3, 100 ms
   "输入_1号梯轿内选层按钮3" : Bool = PLC 输入.1号梯轿内选层按钮3 AT %DB10.DBX2.4, 100 ms
   "输入_1号梯轿内选层按钮4" : Bool = PLC 输入.1号梯轿内选层按钮4 AT %DB10.DBX2.5, 100 ms
   "输入_1号梯轿内选层按钮5" : Bool = PLC 输入.1号梯轿内选层按钮5 AT %DB10.DBX2.6, 100 ms
   "输入_1号梯轿内选层按钮6" : Bool = PLC 输入.1号梯轿内选层按钮6 AT %DB10.DBX2.7, 100 ms
   "输入_1号梯轿内选层按钮7" : Bool = PLC 输入.1号梯轿内选层按钮7 AT %DB10.DBX3.0, 100 ms
   "输入_1号梯轿内选层按钮8" : Bool = PLC 输入.1号梯轿内选层按钮8 AT %DB10.DBX3.1, 100 ms
   "输入_1号梯轿内选层按钮9" : Bool = PLC 输入.1号梯轿内选层按钮9 AT %DB10.DBX3.2, 100 ms
   "输入_1号梯轿内选层按钮10" : Bool = PLC 输入.1号梯轿内选层按钮10 AT %DB10.DBX3.3, 100 ms
   "输出_1号梯LEDa" : Bool = PLC 输出.1号梯LEDa AT %DB11.DBX3.4, 100 ms
   "输出_1号梯LEDb" : Bool = PLC 输出.1号梯LEDb AT %DB11.DBX3.5, 100 ms
   "输出_1号梯LEDc" : Bool = PLC 输出.1号梯LEDc AT %DB11.DBX3.6, 100 ms
   "输出_1号梯LEDd" : Bool = PLC 输出.1号梯LEDd AT %DB11.DBX3.7, 100 ms
   "输出_1号梯LEDe" : Bool = PLC 输出.1号梯LEDe AT %DB11.DBX4.0, 100 ms
   "输出_1号梯LEDf" : Bool = PLC 输出.1号梯LEDf AT %DB11.DBX4.1, 100 ms
   "输出_1号梯LEDi" : Bool = PLC 输出.1号梯LEDi AT %DB11.DBX4.4, 100 ms
   "输出_1号梯LEDj" : Bool = PLC 输出.1号梯LEDj AT %DB11.DBX4.5, 100 ms
   "输出_1号梯1层按钮指示灯" : Bool = PLC 输出.1号梯1层按钮指示灯 AT %DB11.DBX2.2, 100 ms
   "输出_2层上行呼梯按钮指示灯" : Bool = PLC 输出.2层上行呼梯按钮指示灯 AT %DB11.DBX0.1, 100 ms
   "输出_2层下行呼梯按钮指示灯" : Bool = PLC 输出.2层下行呼梯按钮指示灯 AT %DB11.DBX1.1, 100 ms
   "输出_3层上行呼梯按钮指示灯" : Bool = PLC 输出.3层上行呼梯按钮指示灯 AT %DB11.DBX0.2, 100 ms
   "输出_3层下行呼梯按钮指示灯" : Bool = PLC 输出.3层下行呼梯按钮指示灯 AT %DB11.DBX1.2, 100 ms
   "输出_4层上行呼梯按钮指示灯" : Bool = PLC 输出.4层上行呼梯按钮指示灯 AT %DB11.DBX0.3, 100 ms
   "输出_4层下行呼梯按钮指示灯" : Bool = PLC 输出.4层下行呼梯按钮指示灯 AT %DB11.DBX1.3, 100 ms
   "输出_5层上行呼梯按钮指示灯" : Bool = PLC 输出.5层上行呼梯按钮指示灯 AT %DB11.DBX0.4, 100 ms
   "输出_5层下行呼梯按钮指示灯" : Bool = PLC 输出.5层下行呼梯按钮指示灯 AT %DB11.DBX1.4, 100 ms
   "输出_6层上行呼梯按钮指示灯" : Bool = PLC 输出.6层上行呼梯按钮指示灯 AT %DB11.DBX0.5, 100 ms
   "输出_6层下行呼梯按钮指示灯" : Bool = PLC 输出.6层下行呼梯按钮指示灯 AT %DB11.DBX1.5, 100 ms
   "输出_7层上行呼梯按钮指示灯" : Bool = PLC 输出.7层上行呼梯按钮指示灯 AT %DB11.DBX0.6, 100 ms
   "输出_7层下行呼梯按钮指示灯" : Bool = PLC 输出.7层下行呼梯按钮指示灯 AT %DB11.DBX1.6, 100 ms
   "输出_8层上行呼梯按钮指示灯" : Bool = PLC 输出.8层上行呼梯按钮指示灯 AT %DB11.DBX0.7, 100 ms
   "输出_8层下行呼梯按钮指示灯" : Bool = PLC 输出.8层下行呼梯按钮指示灯 AT %DB11.DBX1.7, 100 ms
   "输出_9层上行呼梯按钮指示灯" : Bool = PLC 输出.9层上行呼梯按钮指示灯 AT %DB11.DBX1.0, 100 ms
   "输出_9层下行呼梯按钮指示灯" : Bool = PLC 输出.9层下行呼梯按钮指示灯 AT %DB11.DBX2.0, 100 ms
   "输出_10层下行呼梯按钮指示灯" : Bool = PLC 输出.10层下行呼梯按钮指示灯 AT %DB11.DBX2.1, 100 ms
   "输出_1号梯电机启动信号" : Bool = PLC 输出.1号梯电机启动信号 AT %DB11.DBX6.0, 100 ms
   "输出_1号梯上行接触器" : Bool = PLC 输出.1号梯上行接触器 AT %DB11.DBX6.1, 100 ms
   "输出_1号梯下行接触器" : Bool = PLC 输出.1号梯下行接触器 AT %DB11.DBX6.2, 100 ms
   "输出_1号梯开门继电器" : Bool = PLC 输出.1号梯开门继电器 AT %DB11.DBX6.5, 100 ms
   "输出_1号梯关门继电器" : Bool = PLC 输出.1号梯关门继电器 AT %DB11.DBX6.6, 100 ms
   "输入_1号梯开门到位" : Bool = PLC 输入.1号梯开门到位 AT %DB10.DBX5.3, 100 ms
   "输入_1号梯关门到位" : Bool = PLC 输入.1号梯关门到位 AT %DB10.DBX5.4, 100 ms
   "输出_1号梯低速接触器" : Bool = PLC 输出.1号梯低速接触器 AT %DB11.DBX6.4, 100 ms
   "输出_1号梯高速接触器" : Bool = PLC 输出.1号梯高速接触器 AT %DB11.DBX6.3, 100 ms
   "输出_1号梯1级减速制动" : Bool = PLC 输出.1号梯1级减速制动 AT %DB11.DBX6.7, 100 ms
   "输出_1号梯2级减速制动" : Bool = PLC 输出.1号梯2级减速制动 AT %DB11.DBX7.0, 100 ms
   "输出_1号梯3级减速制动" : Bool = PLC 输出.1号梯3级减速制动 AT %DB11.DBX7.1, 100 ms
   "输入_1号梯检修信号" : Bool = PLC 输入.1号梯检修信号 AT %DB10.DBX3.7, 100 ms
   "输入_1号梯光幕信号" : Bool = PLC 输入.1号梯光幕信号 AT %DB10.DBX3.6, 100 ms
   "输入_1号梯10楼层门锁信号" : Bool = PLC 输入.1号梯10楼层门锁信号 AT %DB10.DBX5.2, 100 ms
   "输入_1号梯9楼层门锁信号" : Bool = PLC 输入.1号梯9楼层门锁信号 AT %DB10.DBX5.1, 100 ms
   "输入_1号梯8楼层门锁信号" : Bool = PLC 输入.1号梯8楼层门锁信号 AT %DB10.DBX5.0, 100 ms
   "输入_1号梯7楼层门锁信号" : Bool = PLC 输入.1号梯7楼层门锁信号 AT %DB10.DBX4.7, 100 ms
   "输入_1号梯6楼层门锁信号" : Bool = PLC 输入.1号梯6楼层门锁信号 AT %DB10.DBX4.6, 100 ms
   "输入_1号梯5楼层门锁信号" : Bool = PLC 输入.1号梯5楼层门锁信号 AT %DB10.DBX4.5, 100 ms
   "输入_1号梯4楼层门锁信号" : Bool = PLC 输入.1号梯4楼层门锁信号 AT %DB10.DBX4.4, 100 ms
   "输入_1号梯3楼层门锁信号" : Bool = PLC 输入.1号梯3楼层门锁信号 AT %DB10.DBX4.3, 100 ms
   "输入_1号梯2楼层门锁信号" : Bool = PLC 输入.1号梯2楼层门锁信号 AT %DB10.DBX4.2, 100 ms
   "输入_1号梯1楼层门锁信号" : Bool = PLC 输入.1号梯1楼层门锁信号 AT %DB10.DBX4.1, 100 ms
   "输入_1号梯轿厢门锁信号" : Bool = PLC 输入.1号梯轿厢门锁信号 AT %DB10.DBX4.0, 100 ms
   "输入_1号梯上端站第2限位" : Bool = PLC 输入.1号梯上端站第2限位 AT %DB10.DBX6.0, 100 ms
   "输入_1号梯上端站第1限位" : Bool = PLC 输入.1号梯上端站第1限位 AT %DB10.DBX5.7, 100 ms
   "输入_1号梯上平层信号" : Bool = PLC 输入.1号梯上平层信号 AT %DB10.DBX5.5, 100 ms
   "输入_1号梯下平层信号" : Bool = PLC 输入.1号梯下平层信号 AT %DB10.DBX5.6, 100 ms
   "输入_1号梯下端站第2限位" : Bool = PLC 输入.1号梯下端站第2限位 AT %DB10.DBX6.2, 100 ms
   "输入_1号梯下端站第1限位" : Bool = PLC 输入.1号梯下端站第1限位 AT %DB10.DBX6.1, 100 ms
   "输出_1号梯上行指示" : Bool = PLC 输出.1号梯上行指示 AT %DB11.DBX5.2, 100 ms
   "输出_1号梯下行指示" : Bool = PLC 输出.1号梯下行指示 AT %DB11.DBX5.3, 100 ms
   "输入_1号梯轿内开门按钮" : Bool = PLC 输入.1号梯轿内开门按钮 AT %DB10.DBX3.4, 100 ms
   "输入_1号梯轿内关门按钮" : Bool = PLC 输入.1号梯轿内关门按钮 AT %DB10.DBX3.5, 100 ms
   "输入_2层下行呼梯按钮" : Bool = PLC 输入.2层下行呼梯按钮 AT %DB10.DBX1.1, 100 ms
   "输出_2号梯满载指示" : Bool = PLC 输出.2号梯满载指示 AT %DB11.DBX10.7, 100 ms
   "输出_2号梯故障指示" : Bool = PLC 输出.2号梯故障指示 AT %DB11.DBX10.4, 100 ms
   "输出_2号梯照明指示" : Bool = PLC 输出.2号梯照明指示 AT %DB11.DBX10.5, 100 ms
   "输出_2号梯风扇指示" : Bool = PLC 输出.2号梯风扇指示 AT %DB11.DBX10.6, 100 ms
   "输出_2号梯上行指示" : Bool = PLC 输出.2号梯上行指示 AT %DB11.DBX10.2, 100 ms
   "输出_2号梯下行指示" : Bool = PLC 输出.2号梯下行指示 AT %DB11.DBX10.3, 100 ms
   "输出_2号梯LEDa" : Bool = PLC 输出.2号梯LEDa AT %DB11.DBX8.4, 100 ms
   "输出_2号梯LEDb" : Bool = PLC 输出.2号梯LEDb AT %DB11.DBX8.5, 100 ms
   "输出_2号梯LEDc" : Bool = PLC 输出.2号梯LEDc AT %DB11.DBX8.6, 100 ms
   "输出_2号梯LEDd" : Bool = PLC 输出.2号梯LEDd AT %DB11.DBX8.7, 100 ms
   "输出_2号梯LEDe" : Bool = PLC 输出.2号梯LEDe AT %DB11.DBX9.0, 100 ms
   "输出_2号梯LEDf" : Bool = PLC 输出.2号梯LEDf AT %DB11.DBX9.1, 100 ms
   "输出_2号梯LEDg" : Bool = PLC 输出.2号梯LEDg AT %DB11.DBX9.2, 100 ms
   "输出_2号梯LEDi" : Bool = PLC 输出.2号梯LEDi AT %DB11.DBX9.4, 100 ms
   "输出_2号梯LEDj" : Bool = PLC 输出.2号梯LEDj AT %DB11.DBX9.5, 100 ms
   "输入_2号梯轿内选层按钮1" : Bool = PLC 输入.2号梯轿内选层按钮1 AT %DB10.DBX6.3, 100 ms
   "输入_2号梯轿内选层按钮2" : Bool = PLC 输入.2号梯轿内选层按钮2 AT %DB10.DBX6.4, 100 ms
   "输入_2号梯轿内选层按钮3" : Bool = PLC 输入.2号梯轿内选层按钮3 AT %DB10.DBX6.5, 100 ms
   "输入_2号梯轿内选层按钮4" : Bool = PLC 输入.2号梯轿内选层按钮4 AT %DB10.DBX6.6, 100 ms
   "输入_2号梯轿内选层按钮5" : Bool = PLC 输入.2号梯轿内选层按钮5 AT %DB10.DBX6.7, 100 ms
   "输入_2号梯轿内选层按钮6" : Bool = PLC 输入.2号梯轿内选层按钮6 AT %DB10.DBX7.0, 100 ms
   "输入_2号梯轿内选层按钮7" : Bool = PLC 输入.2号梯轿内选层按钮7 AT %DB10.DBX7.1, 100 ms
   "输入_2号梯轿内选层按钮8" : Bool = PLC 输入.2号梯轿内选层按钮8 AT %DB10.DBX7.2, 100 ms
   "输入_2号梯轿内选层按钮9" : Bool = PLC 输入.2号梯轿内选层按钮9 AT %DB10.DBX7.3, 100 ms
   "输入_2号梯轿内选层按钮10" : Bool = PLC 输入.2号梯轿内选层按钮10 AT %DB10.DBX7.4, 100 ms
   "输出_2号梯电机启动信号" : Bool = PLC 输出.2号梯电机启动信号 AT %DB11.DBX11.0, 100 ms
   "输出_2号梯上行接触器" : Bool = PLC 输出.2号梯上行接触器 AT %DB11.DBX11.1, 100 ms
   "输出_2号梯下行接触器" : Bool = PLC 输出.2号梯下行接触器 AT %DB11.DBX11.2, 100 ms
   "输出_2号梯开门继电器" : Bool = PLC 输出.2号梯开门继电器 AT %DB11.DBX11.5, 100 ms
   "输出_2号梯关门继电器" : Bool = PLC 输出.2号梯关门继电器 AT %DB11.DBX11.6, 100 ms
   "输入_2号梯开门到位" : Bool = PLC 输入.2号梯开门到位 AT %DB10.DBX9.4, 100 ms
   "输入_2号梯轿内开门按钮" : Bool = PLC 输入.2号梯轿内开门按钮 AT %DB10.DBX7.5, 100 ms
   "输入_2号梯轿内关门按钮" : Bool = PLC 输入.2号梯轿内关门按钮 AT %DB10.DBX7.6, 100 ms
   "输入_2号梯关门到位" : Bool = PLC 输入.2号梯关门到位 AT %DB10.DBX9.5, 100 ms
   "输出_2号梯低速接触器" : Bool = PLC 输出.2号梯低速接触器 AT %DB11.DBX11.4, 100 ms
   "输出_2号梯高速接触器" : Bool = PLC 输出.2号梯高速接触器 AT %DB11.DBX11.3, 100 ms
   "输出_2号梯1级减速制动" : Bool = PLC 输出.2号梯1级减速制动 AT %DB11.DBX11.7, 100 ms
   "输出_2号梯2级减速制动" : Bool = PLC 输出.2号梯2级减速制动 AT %DB11.DBX12.0, 100 ms
   "输出_2号梯3级减速制动" : Bool = PLC 输出.2号梯3级减速制动 AT %DB11.DBX12.1, 100 ms
   "输入_2号梯检修信号" : Bool = PLC 输入.2号梯检修信号 AT %DB10.DBX8.0, 100 ms
   "输入_2号梯光幕信号" : Bool = PLC 输入.2号梯光幕信号 AT %DB10.DBX7.7, 100 ms
   "输入_2号梯10楼层门锁信号" : Bool = PLC 输入.2号梯10楼层门锁信号 AT %DB10.DBX9.3, 100 ms
   "输入_2号梯9楼层门锁信号" : Bool = PLC 输入.2号梯9楼层门锁信号 AT %DB10.DBX9.2, 100 ms
   "输入_2号梯8楼层门锁信号" : Bool = PLC 输入.2号梯8楼层门锁信号 AT %DB10.DBX9.1, 100 ms
   "输入_2号梯7楼层门锁信号" : Bool = PLC 输入.2号梯7楼层门锁信号 AT %DB10.DBX9.0, 100 ms
   "输入_2号梯6楼层门锁信号" : Bool = PLC 输入.2号梯6楼层门锁信号 AT %DB10.DBX8.7, 100 ms
   "输入_2号梯5楼层门锁信号" : Bool = PLC 输入.2号梯5楼层门锁信号 AT %DB10.DBX8.6, 100 ms
   "输入_2号梯4楼层门锁信号" : Bool = PLC 输入.2号梯4楼层门锁信号 AT %DB10.DBX8.5, 100 ms
   "输入_2号梯3楼层门锁信号" : Bool = PLC 输入.2号梯3楼层门锁信号 AT %DB10.DBX8.4, 100 ms
   "输入_2号梯2楼层门锁信号" : Bool = PLC 输入.2号梯2楼层门锁信号 AT %DB10.DBX8.3, 100 ms
   "输入_2号梯1楼层门锁信号" : Bool = PLC 输入.2号梯1楼层门锁信号 AT %DB10.DBX8.2, 100 ms
   "输入_2号梯轿厢门锁信号" : Bool = PLC 输入.2号梯轿厢门锁信号 AT %DB10.DBX8.1, 100 ms
   "输入_2号梯上端站第2限位" : Bool = PLC 输入.2号梯上端站第2限位 AT %DB10.DBX10.1, 100 ms
   "输入_2号梯上端站第1限位" : Bool = PLC 输入.2号梯上端站第1限位 AT %DB10.DBX10.0, 100 ms
   "输入_2号梯下端站第2限位" : Bool = PLC 输入.2号梯下端站第2限位 AT %DB10.DBX10.3, 100 ms
   "输入_3号梯上端站第1限位" : Bool = PLC 输入.3号梯上端站第1限位 AT %DB10.DBX14.1, 100 ms
   "输入_2号梯上平层信号" : Bool = PLC 输入.2号梯上平层信号 AT %DB10.DBX9.6, 100 ms
   "输入_2号梯下平层信号" : Bool = PLC 输入.2号梯下平层信号 AT %DB10.DBX9.7, 100 ms
   "输出_3号梯满载指示" : Bool = PLC 输出.3号梯满载指示 AT %DB11.DBX15.7, 100 ms
   "输出_3号梯故障指示" : Bool = PLC 输出.3号梯故障指示 AT %DB11.DBX15.4, 100 ms
   "输出_3号梯照明指示" : Bool = PLC 输出.3号梯照明指示 AT %DB11.DBX15.5, 100 ms
   "输出_3号梯风扇指示" : Bool = PLC 输出.3号梯风扇指示 AT %DB11.DBX15.6, 100 ms
   "输出_3号梯上行指示" : Bool = PLC 输出.3号梯上行指示 AT %DB11.DBX15.2, 100 ms
   "输出_3号梯下行指示" : Bool = PLC 输出.3号梯下行指示 AT %DB11.DBX15.3, 100 ms
   "输出_3号梯LEDa" : Bool = PLC 输出.3号梯LEDa AT %DB11.DBX13.4, 100 ms
   "输出_3号梯LEDb" : Bool = PLC 输出.3号梯LEDb AT %DB11.DBX13.5, 100 ms
   "输出_3号梯LEDc" : Bool = PLC 输出.3号梯LEDc AT %DB11.DBX13.6, 100 ms
   "输出_3号梯LEDd" : Bool = PLC 输出.3号梯LEDd AT %DB11.DBX13.7, 100 ms
   "输出_3号梯LEDe" : Bool = PLC 输出.3号梯LEDe AT %DB11.DBX14.0, 100 ms
   "输出_3号梯LEDf" : Bool = PLC 输出.3号梯LEDf AT %DB11.DBX14.1, 100 ms
   "输出_3号梯LEDg" : Bool = PLC 输出.3号梯LEDg AT %DB11.DBX14.2, 100 ms
   "输出_3号梯LEDi" : Bool = PLC 输出.3号梯LEDi AT %DB11.DBX14.4, 100 ms
   "输出_3号梯LEDj" : Bool = PLC 输出.3号梯LEDj AT %DB11.DBX14.5, 100 ms
   "输入_3号梯轿内选层按钮10" : Bool = PLC 输入.3号梯轿内选层按钮10 AT %DB10.DBX11.5, 100 ms
   "输入_3号梯轿内选层按钮1" : Bool = PLC 输入.3号梯轿内选层按钮1 AT %DB10.DBX10.4, 100 ms
   "输入_3号梯轿内选层按钮2" : Bool = PLC 输入.3号梯轿内选层按钮2 AT %DB10.DBX10.5, 100 ms
   "输入_3号梯轿内选层按钮3" : Bool = PLC 输入.3号梯轿内选层按钮3 AT %DB10.DBX10.6, 100 ms
   "输入_3号梯轿内选层按钮4" : Bool = PLC 输入.3号梯轿内选层按钮4 AT %DB10.DBX10.7, 100 ms
   "输入_3号梯轿内选层按钮5" : Bool = PLC 输入.3号梯轿内选层按钮5 AT %DB10.DBX11.0, 100 ms
   "输入_3号梯轿内选层按钮6" : Bool = PLC 输入.3号梯轿内选层按钮6 AT %DB10.DBX11.1, 100 ms
   "输入_3号梯轿内选层按钮7" : Bool = PLC 输入.3号梯轿内选层按钮7 AT %DB10.DBX11.2, 100 ms
   "输入_3号梯轿内选层按钮8" : Bool = PLC 输入.3号梯轿内选层按钮8 AT %DB10.DBX11.3, 100 ms
   "输入_3号梯轿内选层按钮9" : Bool = PLC 输入.3号梯轿内选层按钮9 AT %DB10.DBX11.4, 100 ms
   "输出_1层上行呼梯按钮指示灯" : Bool = PLC 输出.1层上行呼梯按钮指示灯 AT %DB11.DBX0.0, 100 ms
   "输出_3号梯电机启动信号" : Bool = PLC 输出.3号梯电机启动信号 AT %DB11.DBX16.0, 100 ms
   "输入_2号梯下端站第1限位" : Bool = PLC 输入.2号梯下端站第1限位 AT %DB10.DBX10.2, 100 ms
   "输出_3号梯上行接触器" : Bool = PLC 输出.3号梯上行接触器 AT %DB11.DBX16.1, 100 ms
   "输出_3号梯下行接触器" : Bool = PLC 输出.3号梯下行接触器 AT %DB11.DBX16.2, 100 ms
   "输出_3号梯开门继电器" : Bool = PLC 输出.3号梯开门继电器 AT %DB11.DBX16.5, 100 ms
   "输出_3号梯关门继电器" : Bool = PLC 输出.3号梯关门继电器 AT %DB11.DBX16.6, 100 ms
   "输入_3号梯开门到位" : Bool = PLC 输入.3号梯开门到位 AT %DB10.DBX13.5, 100 ms
   "输入_3号梯关门到位" : Bool = PLC 输入.3号梯关门到位 AT %DB10.DBX13.6, 100 ms
   "输出_3号梯低速接触器" : Bool = PLC 输出.3号梯低速接触器 AT %DB11.DBX16.4, 100 ms
   "输出_3号梯高速接触器" : Bool = PLC 输出.3号梯高速接触器 AT %DB11.DBX16.3, 100 ms
   "输出_3号梯1级减速制动" : Bool = PLC 输出.3号梯1级减速制动 AT %DB11.DBX16.7, 100 ms
   "输出_3号梯2级减速制动" : Bool = PLC 输出.3号梯2级减速制动 AT %DB11.DBX17.0, 100 ms
   "输出_3号梯3级减速制动" : Bool = PLC 输出.3号梯3级减速制动 AT %DB11.DBX17.1, 100 ms
   "输入_3号梯检修信号" : Bool = PLC 输入.3号梯检修信号 AT %DB10.DBX12.1, 100 ms
   "输入_3号梯光幕信号" : Bool = PLC 输入.3号梯光幕信号 AT %DB10.DBX12.0, 100 ms
   "输入_3号梯10楼层门锁信号" : Bool = PLC 输入.3号梯10楼层门锁信号 AT %DB10.DBX13.4, 100 ms
   "输入_3号梯1楼层门锁信号" : Bool = PLC 输入.3号梯1楼层门锁信号 AT %DB10.DBX12.3, 100 ms
   "输入_3号梯轿厢门锁信号" : Bool = PLC 输入.3号梯轿厢门锁信号 AT %DB10.DBX12.2, 100 ms
   "输入_3号梯2楼层门锁信号" : Bool = PLC 输入.3号梯2楼层门锁信号 AT %DB10.DBX12.4, 100 ms
   "输入_3号梯3楼层门锁信号" : Bool = PLC 输入.3号梯3楼层门锁信号 AT %DB10.DBX12.5, 100 ms
   "输入_3号梯4楼层门锁信号" : Bool = PLC 输入.3号梯4楼层门锁信号 AT %DB10.DBX12.6, 100 ms
   "输入_3号梯5楼层门锁信号" : Bool = PLC 输入.3号梯5楼层门锁信号 AT %DB10.DBX12.7, 100 ms
   "输入_3号梯6楼层门锁信号" : Bool = PLC 输入.3号梯6楼层门锁信号 AT %DB10.DBX13.0, 100 ms
   "输入_3号梯7楼层门锁信号" : Bool = PLC 输入.3号梯7楼层门锁信号 AT %DB10.DBX13.1, 100 ms
   "输入_3号梯8楼层门锁信号" : Bool = PLC 输入.3号梯8楼层门锁信号 AT %DB10.DBX13.2, 100 ms
   "输入_3号梯9楼层门锁信号" : Bool = PLC 输入.3号梯9楼层门锁信号 AT %DB10.DBX13.3, 100 ms
   "输入_3号梯上端站第2限位" : Bool = PLC 输入.3号梯上端站第2限位 AT %DB10.DBX14.2, 100 ms
   "输入_3号梯下端站第2限位" : Bool = PLC 输入.3号梯下端站第2限位 AT %DB10.DBX14.4, 100 ms
   "输入_3号梯下端站第1限位" : Bool = PLC 输入.3号梯下端站第1限位 AT %DB10.DBX14.3, 100 ms
   "输入_3号梯上平层信号" : Bool = PLC 输入.3号梯上平层信号 AT %DB10.DBX13.7, 100 ms
   "输入_3号梯下平层信号" : Bool = PLC 输入.3号梯下平层信号 AT %DB10.DBX14.0, 100 ms
   "输出_4号梯满载指示" : Bool = PLC 输出.4号梯满载指示 AT %DB11.DBX20.7, 100 ms
   "输出_4号梯故障指示" : Bool = PLC 输出.4号梯故障指示 AT %DB11.DBX20.4, 100 ms
   "输出_4号梯照明指示" : Bool = PLC 输出.4号梯照明指示 AT %DB11.DBX20.5, 100 ms
   "输出_4号梯风扇指示" : Bool = PLC 输出.4号梯风扇指示 AT %DB11.DBX20.6, 100 ms
   "输出_4号梯上行指示" : Bool = PLC 输出.4号梯上行指示 AT %DB11.DBX20.2, 100 ms
   "输出_4号梯下行指示" : Bool = PLC 输出.4号梯下行指示 AT %DB11.DBX20.3, 100 ms
   "输出_4号梯LEDa" : Bool = PLC 输出.4号梯LEDa AT %DB11.DBX18.4, 100 ms
   "输出_4号梯LEDb" : Bool = PLC 输出.4号梯LEDb AT %DB11.DBX18.5, 100 ms
   "输出_4号梯LEDc" : Bool = PLC 输出.4号梯LEDc AT %DB11.DBX18.6, 100 ms
   "输出_4号梯LEDd" : Bool = PLC 输出.4号梯LEDd AT %DB11.DBX18.7, 100 ms
   "输出_4号梯LEDe" : Bool = PLC 输出.4号梯LEDe AT %DB11.DBX19.0, 100 ms
   "输出_4号梯LEDf" : Bool = PLC 输出.4号梯LEDf AT %DB11.DBX19.1, 100 ms
   "输出_4号梯LEDg" : Bool = PLC 输出.4号梯LEDg AT %DB11.DBX19.2, 100 ms
   "输出_4号梯LEDi" : Bool = PLC 输出.4号梯LEDi AT %DB11.DBX19.4, 100 ms
   "输出_4号梯LEDj" : Bool = PLC 输出.4号梯LEDj AT %DB11.DBX19.5, 100 ms
   "输出_4号梯电机启动信号" : Bool = PLC 输出.4号梯电机启动信号 AT %DB11.DBX21.0, 100 ms
   "输出_4号梯上行接触器" : Bool = PLC 输出.4号梯上行接触器 AT %DB11.DBX21.1, 100 ms
   "输出_4号梯下行接触器" : Bool = PLC 输出.4号梯下行接触器 AT %DB11.DBX21.2, 100 ms
   "输出_4号梯开门继电器" : Bool = PLC 输出.4号梯开门继电器 AT %DB11.DBX21.5, 100 ms
   "输出_4号梯关门继电器" : Bool = PLC 输出.4号梯关门继电器 AT %DB11.DBX21.6, 100 ms
   "输入_4号梯开门到位" : Bool = PLC 输入.4号梯开门到位 AT %DB10.DBX17.6, 100 ms
   "输入_4号梯关门到位" : Bool = PLC 输入.4号梯关门到位 AT %DB10.DBX17.7, 100 ms
   "输出_4号梯低速接触器" : Bool = PLC 输出.4号梯低速接触器 AT %DB11.DBX21.4, 100 ms
   "输出_4号梯高速接触器" : Bool = PLC 输出.4号梯高速接触器 AT %DB11.DBX21.3, 100 ms
   "输出_4号梯1级减速制动" : Bool = PLC 输出.4号梯1级减速制动 AT %DB11.DBX21.7, 100 ms
   "输出_4号梯2级减速制动" : Bool = PLC 输出.4号梯2级减速制动 AT %DB11.DBX22.0, 100 ms
   "输出_4号梯3级减速制动" : Bool = PLC 输出.4号梯3级减速制动 AT %DB11.DBX22.1, 100 ms
   "输入_4号梯检修信号" : Bool = PLC 输入.4号梯检修信号 AT %DB10.DBX16.2, 100 ms
   "输入_4号梯光幕信号" : Bool = PLC 输入.4号梯光幕信号 AT %DB10.DBX16.1, 100 ms
   "输入_4号梯轿厢门锁信号" : Bool = PLC 输入.4号梯轿厢门锁信号 AT %DB10.DBX16.3, 100 ms
   "输入_4号梯1楼层门锁信号" : Bool = PLC 输入.4号梯1楼层门锁信号 AT %DB10.DBX16.4, 100 ms
   "输入_4号梯2楼层门锁信号" : Bool = PLC 输入.4号梯2楼层门锁信号 AT %DB10.DBX16.5, 100 ms
   "输入_4号梯3楼层门锁信号" : Bool = PLC 输入.4号梯3楼层门锁信号 AT %DB10.DBX16.6, 100 ms
   "输入_4号梯4楼层门锁信号" : Bool = PLC 输入.4号梯4楼层门锁信号 AT %DB10.DBX16.7, 100 ms
   "输入_4号梯5楼层门锁信号" : Bool = PLC 输入.4号梯5楼层门锁信号 AT %DB10.DBX17.0, 100 ms
   "输入_4号梯6楼层门锁信号" : Bool = PLC 输入.4号梯6楼层门锁信号 AT %DB10.DBX17.1, 100 ms
   "输入_4号梯7楼层门锁信号" : Bool = PLC 输入.4号梯7楼层门锁信号 AT %DB10.DBX17.2, 100 ms
   "输入_4号梯8楼层门锁信号" : Bool = PLC 输入.4号梯8楼层门锁信号 AT %DB10.DBX17.3, 100 ms
   "输入_4号梯9楼层门锁信号" : Bool = PLC 输入.4号梯9楼层门锁信号 AT %DB10.DBX17.4, 100 ms
   "输入_4号梯10楼层门锁信号" : Bool = PLC 输入.4号梯10楼层门锁信号 AT %DB10.DBX17.5, 100 ms
   "输入_4号梯上端站第2限位" : Bool = PLC 输入.4号梯上端站第2限位 AT %DB10.DBX18.3, 100 ms
   "输入_4号梯上端站第1限位" : Bool = PLC 输入.4号梯上端站第1限位 AT %DB10.DBX18.2, 100 ms
   "输入_4号梯下平层信号" : Bool = PLC 输入.4号梯下平层信号 AT %DB10.DBX18.1, 100 ms
   "输入_4号梯上平层信号" : Bool = PLC 输入.4号梯上平层信号 AT %DB10.DBX18.0, 100 ms
   "输入_4号梯下端站第2限位" : Bool = PLC 输入.4号梯下端站第2限位 AT %DB10.DBX18.5, 100 ms
   "输入_4号梯下端站第1限位" : Bool = PLC 输入.4号梯下端站第1限位 AT %DB10.DBX18.4, 100 ms
   "输出_1号梯2层按钮指示灯" : Bool = PLC 输出.1号梯2层按钮指示灯 AT %DB11.DBX2.3, 100 ms
   "输出_1号梯3层按钮指示灯" : Bool = PLC 输出.1号梯3层按钮指示灯 AT %DB11.DBX2.4, 100 ms
   "输出_1号梯4层按钮指示灯" : Bool = PLC 输出.1号梯4层按钮指示灯 AT %DB11.DBX2.5, 100 ms
   "输出_1号梯5层按钮指示灯" : Bool = PLC 输出.1号梯5层按钮指示灯 AT %DB11.DBX2.6, 100 ms
   "输出_1号梯6层按钮指示灯" : Bool = PLC 输出.1号梯6层按钮指示灯 AT %DB11.DBX2.7, 100 ms
   "输出_1号梯7层按钮指示灯" : Bool = PLC 输出.1号梯7层按钮指示灯 AT %DB11.DBX3.0, 100 ms
   "输出_1号梯8层按钮指示灯" : Bool = PLC 输出.1号梯8层按钮指示灯 AT %DB11.DBX3.1, 100 ms
   "输出_1号梯9层按钮指示灯" : Bool = PLC 输出.1号梯9层按钮指示灯 AT %DB11.DBX3.2, 100 ms
   "输出_1号梯10层按钮指示灯" : Bool = PLC 输出.1号梯10层按钮指示灯 AT %DB11.DBX3.3, 100 ms
   "输出_2号梯10层按钮指示灯" : Bool = PLC 输出.2号梯10层按钮指示灯 AT %DB11.DBX8.3, 100 ms
   "输出_2号梯9层按钮指示灯" : Bool = PLC 输出.2号梯9层按钮指示灯 AT %DB11.DBX8.2, 100 ms
   "输出_2号梯8层按钮指示灯" : Bool = PLC 输出.2号梯8层按钮指示灯 AT %DB11.DBX8.1, 100 ms
   "输出_2号梯7层按钮指示灯" : Bool = PLC 输出.2号梯7层按钮指示灯 AT %DB11.DBX8.0, 100 ms
   "输出_2号梯6层按钮指示灯" : Bool = PLC 输出.2号梯6层按钮指示灯 AT %DB11.DBX7.7, 100 ms
   "输出_2号梯5层按钮指示灯" : Bool = PLC 输出.2号梯5层按钮指示灯 AT %DB11.DBX7.6, 100 ms
   "输出_2号梯4层按钮指示灯" : Bool = PLC 输出.2号梯4层按钮指示灯 AT %DB11.DBX7.5, 100 ms
   "输出_2号梯3层按钮指示灯" : Bool = PLC 输出.2号梯3层按钮指示灯 AT %DB11.DBX7.4, 100 ms
   "输出_2号梯2层按钮指示灯" : Bool = PLC 输出.2号梯2层按钮指示灯 AT %DB11.DBX7.3, 100 ms
   "输出_2号梯1层按钮指示灯" : Bool = PLC 输出.2号梯1层按钮指示灯 AT %DB11.DBX7.2, 100 ms
   "输出_3号梯1层按钮指示灯" : Bool = PLC 输出.3号梯1层按钮指示灯 AT %DB11.DBX12.2, 100 ms
   "输出_3号梯2层按钮指示灯" : Bool = PLC 输出.3号梯2层按钮指示灯 AT %DB11.DBX12.3, 100 ms
   "输出_3号梯3层按钮指示灯" : Bool = PLC 输出.3号梯3层按钮指示灯 AT %DB11.DBX12.4, 100 ms
   "输出_3号梯4层按钮指示灯" : Bool = PLC 输出.3号梯4层按钮指示灯 AT %DB11.DBX12.5, 100 ms
   "输出_3号梯5层按钮指示灯" : Bool = PLC 输出.3号梯5层按钮指示灯 AT %DB11.DBX12.6, 100 ms
   "输出_3号梯6层按钮指示灯" : Bool = PLC 输出.3号梯6层按钮指示灯 AT %DB11.DBX12.7, 100 ms
   "输出_3号梯7层按钮指示灯" : Bool = PLC 输出.3号梯7层按钮指示灯 AT %DB11.DBX13.0, 100 ms
   "输出_3号梯8层按钮指示灯" : Bool = PLC 输出.3号梯8层按钮指示灯 AT %DB11.DBX13.1, 100 ms
   "输出_3号梯9层按钮指示灯" : Bool = PLC 输出.3号梯9层按钮指示灯 AT %DB11.DBX13.2, 100 ms
   "输出_3号梯10层按钮指示灯" : Bool = PLC 输出.3号梯10层按钮指示灯 AT %DB11.DBX13.3, 100 ms
   "输出_4号梯1层按钮指示灯" : Bool = PLC 输出.4号梯1层按钮指示灯 AT %DB11.DBX17.2, 100 ms
   "输出_4号梯2层按钮指示灯" : Bool = PLC 输出.4号梯2层按钮指示灯 AT %DB11.DBX17.3, 100 ms
   "输出_4号梯3层按钮指示灯" : Bool = PLC 输出.4号梯3层按钮指示灯 AT %DB11.DBX17.4, 100 ms
   "输出_4号梯4层按钮指示灯" : Bool = PLC 输出.4号梯4层按钮指示灯 AT %DB11.DBX17.5, 100 ms
   "输出_4号梯5层按钮指示灯" : Bool = PLC 输出.4号梯5层按钮指示灯 AT %DB11.DBX17.6, 100 ms
   "输出_4号梯6层按钮指示灯" : Bool = PLC 输出.4号梯6层按钮指示灯 AT %DB11.DBX17.7, 100 ms
   "输出_4号梯7层按钮指示灯" : Bool = PLC 输出.4号梯7层按钮指示灯 AT %DB11.DBX18.0, 100 ms
   "输出_4号梯8层按钮指示灯" : Bool = PLC 输出.4号梯8层按钮指示灯 AT %DB11.DBX18.1, 100 ms
   "输出_4号梯9层按钮指示灯" : Bool = PLC 输出.4号梯9层按钮指示灯 AT %DB11.DBX18.2, 100 ms
   "输出_4号梯10层按钮指示灯" : Bool = PLC 输出.4号梯10层按钮指示灯 AT %DB11.DBX18.3, 100 ms
   "输出_5号梯满载指示" : Bool = PLC 输出.5号梯满载指示 AT %DB11.DBX25.7, 100 ms
   "输出_6号梯满载指示" : Bool = PLC 输出.6号梯满载指示 AT %DB11.DBX30.7, 100 ms
   "输出_6号梯故障指示" : Bool = PLC 输出.6号梯故障指示 AT %DB11.DBX30.4, 100 ms
   "输出_5号梯故障指示" : Bool = PLC 输出.5号梯故障指示 AT %DB11.DBX25.4, 100 ms
   "输出_5号梯照明指示" : Bool = PLC 输出.5号梯照明指示 AT %DB11.DBX25.5, 100 ms
   "输出_6号梯照明指示" : Bool = PLC 输出.6号梯照明指示 AT %DB11.DBX30.5, 100 ms
   "输出_6号梯风扇指示" : Bool = PLC 输出.6号梯风扇指示 AT %DB11.DBX30.6, 100 ms
   "输出_5号梯风扇指示" : Bool = PLC 输出.5号梯风扇指示 AT %DB11.DBX25.6, 100 ms
   "输出_5号梯上行指示" : Bool = PLC 输出.5号梯上行指示 AT %DB11.DBX25.2, 100 ms
   "输出_5号梯下行指示" : Bool = PLC 输出.5号梯下行指示 AT %DB11.DBX25.3, 100 ms
   "输出_5号梯LEDa" : Bool = PLC 输出.5号梯LEDa AT %DB11.DBX23.4, 100 ms
   "输出_5号梯LEDb" : Bool = PLC 输出.5号梯LEDb AT %DB11.DBX23.5, 100 ms
   "输出_5号梯LEDc" : Bool = PLC 输出.5号梯LEDc AT %DB11.DBX23.6, 100 ms
   "输出_5号梯LEDd" : Bool = PLC 输出.5号梯LEDd AT %DB11.DBX23.7, 100 ms
   "输出_5号梯LEDe" : Bool = PLC 输出.5号梯LEDe AT %DB11.DBX24.0, 100 ms
   "输出_5号梯LEDf" : Bool = PLC 输出.5号梯LEDf AT %DB11.DBX24.1, 100 ms
   "输出_5号梯LEDg" : Bool = PLC 输出.5号梯LEDg AT %DB11.DBX24.2, 100 ms
   "输出_5号梯LEDi" : Bool = PLC 输出.5号梯LEDi AT %DB11.DBX24.4, 100 ms
   "输出_5号梯LEDj" : Bool = PLC 输出.5号梯LEDj AT %DB11.DBX24.5, 100 ms
   "输入_5号梯轿内开门按钮" : Bool = PLC 输入.5号梯轿内开门按钮 AT %DB10.DBX20.0, 100 ms
   "输入_5号梯轿内关门按钮" : Bool = PLC 输入.5号梯轿内关门按钮 AT %DB10.DBX20.1, 100 ms
   "输入_4号梯轿内开门按钮" : Bool = PLC 输入.4号梯轿内开门按钮 AT %DB10.DBX15.7, 100 ms
   "输入_4号梯轿内关门按钮" : Bool = PLC 输入.4号梯轿内关门按钮 AT %DB10.DBX16.0, 100 ms
   "输入_3号梯轿内开门按钮" : Bool = PLC 输入.3号梯轿内开门按钮 AT %DB10.DBX11.6, 100 ms
   "输入_3号梯轿内关门按钮" : Bool = PLC 输入.3号梯轿内关门按钮 AT %DB10.DBX11.7, 100 ms
   "输入_5号梯轿内选层按钮1" : Bool = PLC 输入.5号梯轿内选层按钮1 AT %DB10.DBX18.6, 100 ms
   "输出_5号梯1层按钮指示灯" : Bool = PLC 输出.5号梯1层按钮指示灯 AT %DB11.DBX22.2, 100 ms
   "输入_5号梯轿内选层按钮2" : Bool = PLC 输入.5号梯轿内选层按钮2 AT %DB10.DBX18.7, 100 ms
   "输出_5号梯3层按钮指示灯" : Bool = PLC 输出.5号梯3层按钮指示灯 AT %DB11.DBX22.4, 100 ms
   "输入_5号梯轿内选层按钮3" : Bool = PLC 输入.5号梯轿内选层按钮3 AT %DB10.DBX19.0, 100 ms
   "输入_5号梯轿内选层按钮4" : Bool = PLC 输入.5号梯轿内选层按钮4 AT %DB10.DBX19.1, 100 ms
   "输入_5号梯轿内选层按钮5" : Bool = PLC 输入.5号梯轿内选层按钮5 AT %DB10.DBX19.2, 100 ms
   "输入_5号梯轿内选层按钮6" : Bool = PLC 输入.5号梯轿内选层按钮6 AT %DB10.DBX19.3, 100 ms
   "输入_5号梯轿内选层按钮7" : Bool = PLC 输入.5号梯轿内选层按钮7 AT %DB10.DBX19.4, 100 ms
   "输入_5号梯轿内选层按钮8" : Bool = PLC 输入.5号梯轿内选层按钮8 AT %DB10.DBX19.5, 100 ms
   "输入_5号梯轿内选层按钮9" : Bool = PLC 输入.5号梯轿内选层按钮9 AT %DB10.DBX19.6, 100 ms
   "输入_5号梯轿内选层按钮10" : Bool = PLC 输入.5号梯轿内选层按钮10 AT %DB10.DBX19.7, 100 ms
   "输出_5号梯10层按钮指示灯" : Bool = PLC 输出.5号梯10层按钮指示灯 AT %DB11.DBX23.3, 100 ms
   "输出_5号梯9层按钮指示灯" : Bool = PLC 输出.5号梯9层按钮指示灯 AT %DB11.DBX23.2, 100 ms
   "输出_5号梯8层按钮指示灯" : Bool = PLC 输出.5号梯8层按钮指示灯 AT %DB11.DBX23.1, 100 ms
   "输出_5号梯7层按钮指示灯" : Bool = PLC 输出.5号梯7层按钮指示灯 AT %DB11.DBX23.0, 100 ms
   "输出_5号梯6层按钮指示灯" : Bool = PLC 输出.5号梯6层按钮指示灯 AT %DB11.DBX22.7, 100 ms
   "输出_5号梯5层按钮指示灯" : Bool = PLC 输出.5号梯5层按钮指示灯 AT %DB11.DBX22.6, 100 ms
   "输出_5号梯4层按钮指示灯" : Bool = PLC 输出.5号梯4层按钮指示灯 AT %DB11.DBX22.5, 100 ms
   "输出_5号梯2层按钮指示灯" : Bool = PLC 输出.5号梯2层按钮指示灯 AT %DB11.DBX22.3, 100 ms
   "输出_5号梯电机启动信号" : Bool = PLC 输出.5号梯电机启动信号 AT %DB11.DBX26.0, 100 ms
   "输出_5号梯上行接触器" : Bool = PLC 输出.5号梯上行接触器 AT %DB11.DBX26.1, 100 ms
   "输出_5号梯下行接触器" : Bool = PLC 输出.5号梯下行接触器 AT %DB11.DBX26.2, 100 ms
   "输出_5号梯开门继电器" : Bool = PLC 输出.5号梯开门继电器 AT %DB11.DBX26.5, 100 ms
   "输出_5号梯关门继电器" : Bool = PLC 输出.5号梯关门继电器 AT %DB11.DBX26.6, 100 ms
   "输入_5号梯开门到位" : Bool = PLC 输入.5号梯开门到位 AT %DB10.DBX21.7, 100 ms
   "输入_5号梯关门到位" : Bool = PLC 输入.5号梯关门到位 AT %DB10.DBX22.0, 100 ms
   "输出_5号梯低速接触器" : Bool = PLC 输出.5号梯低速接触器 AT %DB11.DBX26.4, 100 ms
   "输出_5号梯高速接触器" : Bool = PLC 输出.5号梯高速接触器 AT %DB11.DBX26.3, 100 ms
   "输出_5号梯1级减速制动" : Bool = PLC 输出.5号梯1级减速制动 AT %DB11.DBX26.7, 100 ms
   "输出_5号梯2级减速制动" : Bool = PLC 输出.5号梯2级减速制动 AT %DB11.DBX27.0, 100 ms
   "输出_5号梯3级减速制动" : Bool = PLC 输出.5号梯3级减速制动 AT %DB11.DBX27.1, 100 ms
   "输入_5号梯检修信号" : Bool = PLC 输入.5号梯检修信号 AT %DB10.DBX20.3, 100 ms
   "输入_5号梯光幕信号" : Bool = PLC 输入.5号梯光幕信号 AT %DB10.DBX20.2, 100 ms
   "输入_5号梯10楼层门锁信号" : Bool = PLC 输入.5号梯10楼层门锁信号 AT %DB10.DBX21.6, 100 ms
   "输入_5号梯1楼层门锁信号" : Bool = PLC 输入.5号梯1楼层门锁信号 AT %DB10.DBX20.5, 100 ms
   "输入_5号梯轿厢门锁信号" : Bool = PLC 输入.5号梯轿厢门锁信号 AT %DB10.DBX20.4, 100 ms
   "输入_5号梯2楼层门锁信号" : Bool = PLC 输入.5号梯2楼层门锁信号 AT %DB10.DBX20.6, 100 ms
   "输入_5号梯3楼层门锁信号" : Bool = PLC 输入.5号梯3楼层门锁信号 AT %DB10.DBX20.7, 100 ms
   "输入_5号梯4楼层门锁信号" : Bool = PLC 输入.5号梯4楼层门锁信号 AT %DB10.DBX21.0, 100 ms
   "输入_5号梯6楼层门锁信号" : Bool = PLC 输入.5号梯6楼层门锁信号 AT %DB10.DBX21.2, 100 ms
   "输入_5号梯7楼层门锁信号" : Bool = PLC 输入.5号梯7楼层门锁信号 AT %DB10.DBX21.3, 100 ms
   "输入_5号梯8楼层门锁信号" : Bool = PLC 输入.5号梯8楼层门锁信号 AT %DB10.DBX21.4, 100 ms
   "输入_5号梯9楼层门锁信号" : Bool = PLC 输入.5号梯9楼层门锁信号 AT %DB10.DBX21.5, 100 ms
   "输入_5号梯上端站第2限位" : Bool = PLC 输入.5号梯上端站第2限位 AT %DB10.DBX22.4, 100 ms
   "输入_5号梯上端站第1限位" : Bool = PLC 输入.5号梯上端站第1限位 AT %DB10.DBX22.3, 100 ms
   "输入_5号梯下端站第1限位" : Bool = PLC 输入.5号梯下端站第1限位 AT %DB10.DBX22.5, 100 ms
   "输入_5号梯下端站第2限位" : Bool = PLC 输入.5号梯下端站第2限位 AT %DB10.DBX22.6, 100 ms
   "输入_5号梯上平层信号" : Bool = PLC 输入.5号梯上平层信号 AT %DB10.DBX22.1, 100 ms
   "输入_5号梯下平层信号" : Bool = PLC 输入.5号梯下平层信号 AT %DB10.DBX22.2, 100 ms
   "输出_6号梯上行指示" : Bool = PLC 输出.6号梯上行指示 AT %DB11.DBX30.2, 100 ms
   "输出_6号梯下行指示" : Bool = PLC 输出.6号梯下行指示 AT %DB11.DBX30.3, 100 ms
   "输出_6号梯LEDa" : Bool = PLC 输出.6号梯LEDa AT %DB11.DBX28.4, 100 ms
   "输出_6号梯LEDb" : Bool = PLC 输出.6号梯LEDb AT %DB11.DBX28.5, 100 ms
   "输出_6号梯LEDc" : Bool = PLC 输出.6号梯LEDc AT %DB11.DBX28.6, 100 ms
   "输出_6号梯LEDd" : Bool = PLC 输出.6号梯LEDd AT %DB11.DBX28.7, 100 ms
   "输出_6号梯LEDe" : Bool = PLC 输出.6号梯LEDe AT %DB11.DBX29.0, 100 ms
   "输出_6号梯LEDf" : Bool = PLC 输出.6号梯LEDf AT %DB11.DBX29.1, 100 ms
   "输出_6号梯LEDg" : Bool = PLC 输出.6号梯LEDg AT %DB11.DBX29.2, 100 ms
   "输出_6号梯LEDi" : Bool = PLC 输出.6号梯LEDi AT %DB11.DBX29.4, 100 ms
   "输出_6号梯LEDj" : Bool = PLC 输出.6号梯LEDj AT %DB11.DBX29.5, 100 ms
   "输入_6号梯轿内开门按钮" : Bool = PLC 输入.6号梯轿内开门按钮 AT %DB10.DBX24.1, 100 ms
   "输出_6号梯电机启动信号" : Bool = PLC 输出.6号梯电机启动信号 AT %DB11.DBX31.0, 100 ms
   "输出_6号梯开门继电器" : Bool = PLC 输出.6号梯开门继电器 AT %DB11.DBX31.5, 100 ms
   "输出_6号梯关门继电器" : Bool = PLC 输出.6号梯关门继电器 AT %DB11.DBX31.6, 100 ms
   "输入_6号梯开门到位" : Bool = PLC 输入.6号梯开门到位 AT %DB10.DBX26.0, 100 ms
   "输入_6号梯关门到位" : Bool = PLC 输入.6号梯关门到位 AT %DB10.DBX26.1, 100 ms
   "输出_6号梯低速接触器" : Bool = PLC 输出.6号梯低速接触器 AT %DB11.DBX31.4, 100 ms
   "输出_6号梯高速接触器" : Bool = PLC 输出.6号梯高速接触器 AT %DB11.DBX31.3, 100 ms
   "输出_6号梯1级减速制动" : Bool = PLC 输出.6号梯1级减速制动 AT %DB11.DBX31.7, 100 ms
   "输出_6号梯2级减速制动" : Bool = PLC 输出.6号梯2级减速制动 AT %DB11.DBX32.0, 100 ms
   "输出_6号梯3级减速制动" : Bool = PLC 输出.6号梯3级减速制动 AT %DB11.DBX32.1, 100 ms
   "输入_6号梯检修信号" : Bool = PLC 输入.6号梯检修信号 AT %DB10.DBX24.4, 100 ms
   "输入_6号梯光幕信号" : Bool = PLC 输入.6号梯光幕信号 AT %DB10.DBX24.3, 100 ms
   "输入_6号梯轿厢门锁信号" : Bool = PLC 输入.6号梯轿厢门锁信号 AT %DB10.DBX24.5, 100 ms
   "输入_6号梯1楼层门锁信号" : Bool = PLC 输入.6号梯1楼层门锁信号 AT %DB10.DBX24.6, 100 ms
   "输入_6号梯2楼层门锁信号" : Bool = PLC 输入.6号梯2楼层门锁信号 AT %DB10.DBX24.7, 100 ms
   "输入_6号梯3楼层门锁信号" : Bool = PLC 输入.6号梯3楼层门锁信号 AT %DB10.DBX25.0, 100 ms
   "输入_6号梯4楼层门锁信号" : Bool = PLC 输入.6号梯4楼层门锁信号 AT %DB10.DBX25.1, 100 ms
   "输入_6号梯5楼层门锁信号" : Bool = PLC 输入.6号梯5楼层门锁信号 AT %DB10.DBX25.2, 100 ms
   "输入_6号梯6楼层门锁信号" : Bool = PLC 输入.6号梯6楼层门锁信号 AT %DB10.DBX25.3, 100 ms
   "输入_6号梯8楼层门锁信号" : Bool = PLC 输入.6号梯8楼层门锁信号 AT %DB10.DBX25.5, 100 ms
   "输入_6号梯7楼层门锁信号" : Bool = PLC 输入.6号梯7楼层门锁信号 AT %DB10.DBX25.4, 100 ms
   "输入_6号梯9楼层门锁信号" : Bool = PLC 输入.6号梯9楼层门锁信号 AT %DB10.DBX25.6, 100 ms
   "输入_6号梯10楼层门锁信号" : Bool = PLC 输入.6号梯10楼层门锁信号 AT %DB10.DBX25.7, 100 ms
   "输入_6号梯下端站第1限位" : Bool = PLC 输入.6号梯下端站第1限位 AT %DB10.DBX26.6, 100 ms
   "输入_6号梯下端站第2限位" : Bool = PLC 输入.6号梯下端站第2限位 AT %DB10.DBX26.7, 100 ms
   "输入_6号梯上端站第1限位" : Bool = PLC 输入.6号梯上端站第1限位 AT %DB10.DBX26.4, 100 ms
   "输入_6号梯上端站第2限位" : Bool = PLC 输入.6号梯上端站第2限位 AT %DB10.DBX26.5, 100 ms
   "输入_6号梯上平层信号" : Bool = PLC 输入.6号梯上平层信号 AT %DB10.DBX26.2, 100 ms
   "输入_6号梯下平层信号" : Bool = PLC 输入.6号梯下平层信号 AT %DB10.DBX26.3, 100 ms
   "username" : WString[10], internal
   "zuhao" : UInt, internal
   "1号梯初始化变量" : Int = PLC 中间变量1.1号梯初始化楼层数 AT %DB13.DBW42, 100 ms
   "6号梯初始化变量" : Int = PLC 中间变量1.6号梯初始化楼层数 AT %DB13.DBW52, 100 ms
   "输出_1号梯LEDg" : Bool = PLC 输出.1号梯LEDg AT %DB11.DBX4.2, 100 ms
   "5号梯初始化变量" : Int = PLC 中间变量1.5号梯初始化楼层数 AT %DB13.DBW50, 100 ms
   "4号梯初始化变量" : Int = PLC 中间变量1.4号梯初始化楼层数 AT %DB13.DBW48, 100 ms
   "3号梯初始化变量" : Int = PLC 中间变量1.3号梯初始化楼层数 AT %DB13.DBW46, 100 ms
   "2号梯初始化变量" : Int = PLC 中间变量1.2号梯初始化楼层数 AT %DB13.DBW44, 100 ms
   "输出_6号梯1层按钮指示灯" : Bool = PLC 输出.6号梯1层按钮指示灯 AT %DB11.DBX27.2, 100 ms
   "输出_6号梯2层按钮指示灯" : Bool = PLC 输出.6号梯2层按钮指示灯 AT %DB11.DBX27.3, 100 ms
   "输出_6号梯3层按钮指示灯" : Bool = PLC 输出.6号梯3层按钮指示灯 AT %DB11.DBX27.4, 100 ms
   "输出_6号梯4层按钮指示灯" : Bool = PLC 输出.6号梯4层按钮指示灯 AT %DB11.DBX27.5, 100 ms
   "输出_6号梯5层按钮指示灯" : Bool = PLC 输出.6号梯5层按钮指示灯 AT %DB11.DBX27.6, 100 ms
   "输出_6号梯6层按钮指示灯" : Bool = PLC 输出.6号梯6层按钮指示灯 AT %DB11.DBX27.7, 100 ms
   "输出_6号梯7层按钮指示灯" : Bool = PLC 输出.6号梯7层按钮指示灯 AT %DB11.DBX28.0, 100 ms
   "输出_6号梯8层按钮指示灯" : Bool = PLC 输出.6号梯8层按钮指示灯 AT %DB11.DBX28.1, 100 ms
   "输出_6号梯9层按钮指示灯" : Bool = PLC 输出.6号梯9层按钮指示灯 AT %DB11.DBX28.2, 100 ms
   "输出_6号梯10层按钮指示灯" : Bool = PLC 输出.6号梯10层按钮指示灯 AT %DB11.DBX28.3, 100 ms
   "1号梯正常运行" : Bool = PLC 中间变量1.1号梯准备就绪 AT %DB13.DBX100.0, 100 ms
   "1号梯满载故障" : Bool = PLC 输出.1号梯满载指示 AT %DB11.DBX5.7, 100 ms
   "1号梯检修" : Bool = PLC 输入.1号梯检修信号 AT %DB10.DBX3.7, 100 ms
   "2号梯正常运行" : Bool = PLC 中间变量1.2号梯准备就绪 AT %DB13.DBX100.1, 100 ms
   "3号梯正常运行" : Bool = PLC 中间变量1.3号梯准备就绪 AT %DB13.DBX100.2, 100 ms
   "4号梯正常运行" : Bool = PLC 中间变量1.4号梯准备就绪 AT %DB13.DBX100.3, 100 ms
   "5号梯正常运行" : Bool = PLC 中间变量1.5号梯准备就绪 AT %DB13.DBX100.4, 100 ms
   "6号梯正常运行" : Bool = PLC 中间变量1.6号梯准备就绪 AT %DB13.DBX100.5, 100 ms
   "2号梯满载故障" : Bool = PLC 输出.2号梯满载指示 AT %DB11.DBX10.7, 100 ms
   "3号梯满载故障" : Bool = PLC 输出.3号梯满载指示 AT %DB11.DBX15.7, 100 ms
   "5号梯满载故障" : Bool = PLC 输出.5号梯满载指示 AT %DB11.DBX25.7, 100 ms
   "4号梯满载故障" : Bool = PLC 输出.4号梯满载指示 AT %DB11.DBX20.7, 100 ms
   "6号梯满载故障" : Bool = PLC 输出.6号梯满载指示 AT %DB11.DBX30.7, 100 ms
   "2号梯检修" : Bool = PLC 输入.2号梯检修信号 AT %DB10.DBX8.0, 100 ms
   "3号梯检修" : Bool = PLC 输入.3号梯检修信号 AT %DB10.DBX12.1, 100 ms
   "4号梯检修" : Bool = PLC 输入.4号梯检修信号 AT %DB10.DBX16.2, 100 ms
   "5号梯检修" : Bool = PLC 输入.5号梯检修信号 AT %DB10.DBX20.3, 100 ms
   "6号梯检修" : Bool = PLC 输入.6号梯检修信号 AT %DB10.DBX24.4, 100 ms

HMI tags "默认变量表2"
   "1号电梯初始化终点楼层" : Int = PLC 中间变量1.1号梯初始化楼层数 AT %DB13.DBW42, 100 ms
   "2号电梯初始化终点楼层" : Int = PLC 中间变量1.2号梯初始化楼层数 AT %DB13.DBW44, 100 ms
   "3号电梯初始化终点楼层" : Int = PLC 中间变量1.3号梯初始化楼层数 AT %DB13.DBW46, 100 ms
   "4号电梯初始化终点楼层" : Int = PLC 中间变量1.4号梯初始化楼层数 AT %DB13.DBW48, 100 ms
   "5号电梯初始化终点楼层" : Int = PLC 中间变量1.5号梯初始化楼层数 AT %DB13.DBW50, 100 ms
   "6号电梯初始化终点楼层" : Int = PLC 中间变量1.6号梯初始化楼层数 AT %DB13.DBW52, 100 ms
   "1号电梯电梯初始化方向向上" : Bool = PLC 中间变量1.1号梯初始化方向上行 AT %DB13.DBX54.6, 100 ms
   "2号电梯电梯初始化方向向上" : Bool = PLC 中间变量1.2号梯初始化方向上行 AT %DB13.DBX54.7, 100 ms
   "5号电梯电梯初始化方向向上" : Bool = PLC 中间变量1.5号梯初始化方向上行 AT %DB13.DBX55.2, 100 ms
   "3号电梯电梯初始化方向向上" : Bool = PLC 中间变量1.3号梯初始化方向上行 AT %DB13.DBX55.0, 100 ms
   "4号电梯电梯初始化方向向上" : Bool = PLC 中间变量1.4号梯初始化方向上行 AT %DB13.DBX55.1, 100 ms
   "6号电梯电梯初始化方向向上" : Bool = PLC 中间变量1.6号梯初始化方向上行 AT %DB13.DBX55.3, 100 ms

HMI tags "默认变量表3"
   "初始化设置用_1号梯初始化方向选择" : Int = PLC 中间变量1.1号梯初始化方向位 AT %DB13.DBW118, 100 ms
   "初始化设置用_2号梯初始化方向选择" : Int = PLC 中间变量1.2号梯初始化方向位 AT %DB13.DBW120, 100 ms
   "初始化设置用_3号梯初始化方向选择" : Int = PLC 中间变量1.3号梯初始化方向位 AT %DB13.DBW122, 100 ms
   "初始化设置用_4号梯初始化方向选择" : Int = PLC 中间变量1.4号梯初始化方向位 AT %DB13.DBW124, 100 ms
   "初始化设置用_5号梯初始化方向选择" : Int = PLC 中间变量1.5号梯初始化方向位 AT %DB13.DBW126, 100 ms
   "初始化设置用_6号梯初始化方向选择" : Int = PLC 中间变量1.6号梯初始化方向位 AT %DB13.DBW128, 100 ms
   "初始化设置用_1号梯初始化楼层赋值" : Int = PLC 中间变量1.1号梯初始化楼层数 AT %DB13.DBW42, 100 ms
   "初始化设置用_2号梯初始化楼层赋值" : Int = PLC 中间变量1.2号梯初始化楼层数 AT %DB13.DBW44, 100 ms
   "初始化设置用_3号梯初始化楼层赋值" : Int = PLC 中间变量1.3号梯初始化楼层数 AT %DB13.DBW46, 100 ms
   "初始化设置用_4号梯初始化楼层赋值" : Int = PLC 中间变量1.4号梯初始化楼层数 AT %DB13.DBW48, 100 ms
   "初始化设置用_5号梯初始化楼层赋值" : Int = PLC 中间变量1.5号梯初始化楼层数 AT %DB13.DBW50, 100 ms
   "初始化设置用_6号梯初始化楼层赋值" : Int = PLC 中间变量1.6号梯初始化楼层数 AT %DB13.DBW52, 100 ms
   "1号梯载重量" : Int = PLC 中间变量2.1号梯转换后载重量 AT %DB3.DBW712, 100 ms
   "输入_1号梯当前载重量" : Word = PLC 输入.1号梯当前载重量 AT %DB10.DBW28, 100 ms
   "2号梯载重量" : Int = PLC 中间变量2.2号梯转换后载重量 AT %DB3.DBW714, 100 ms
   "3号梯载重量" : Int = PLC 中间变量2.3号梯转换后载重量 AT %DB3.DBW716, 100 ms
   "4号梯载重量" : Int = PLC 中间变量2.4号梯转换后载重量 AT %DB3.DBW718, 100 ms
   "5号梯载重量" : Int = PLC 中间变量2.5号梯转换后载重量 AT %DB3.DBW720, 100 ms
   "6号梯载重量" : Int = PLC 中间变量2.6号梯转换后载重量 AT %DB3.DBW722, 100 ms
   "输入_2号梯当前载重量" : Word = PLC 输入.2号梯当前载重量 AT %DB10.DBW30, 100 ms
   "输入_3号梯当前载重量" : Word = PLC 输入.3号梯当前载重量 AT %DB10.DBW32, 100 ms
   "输入_4号梯当前载重量" : Word = PLC 输入.4号梯当前载重量 AT %DB10.DBW34, 100 ms
   "输入_5号梯当前载重量" : Word = PLC 输入.5号梯当前载重量 AT %DB10.DBW36, 100 ms
   "输入_6号梯当前载重量" : Word = PLC 输入.6号梯当前载重量 AT %DB10.DBW38, 100 ms
   "程序运行秒" : Int = PLC 中间变量1.程序运行时长秒 AT %DB13.DBW146, 100 ms
   "程序运行分钟" : Int = PLC 中间变量1.程序运行时长分钟 AT %DB13.DBW148, 100 ms
   "程序运行小时" : Int = PLC 中间变量1.程序运行时长小时 AT %DB13.DBW150, 100 ms

text list "zuhao": 1 '管理员'; 2 '监视员'; 3 '操作员'

text list "身份": 1 '监视员'; 0 '操作员'; 0 '管理员'

recipe "配方1": 1号梯上端站第1限位 <- "输入_1号梯上端站第1限位", 1号梯上端站第2限位 <- "输入_1号梯上端站第2限位", 1号梯下端站第1限位 <- "输入_1号梯下端站第1限位", 1号梯下端站第2限位 <- "输入_1号梯下端站第2限位", 2号梯上端站第1限位 <- "输入_2号梯上端站第1限位", 2号梯上端站第2限位 <- "输入_2号梯上端站第2限位", 2号梯下端站第1限位 <- "输入_2号梯下端站第1限位", 2号梯下端站第2限位 <- "输入_2号梯下端站第2限位", 3号梯上端站第1限位 <- "输入_3号梯上端站第1限位", 3号梯上端站第2限位 <- "输入_3号梯上端站第2限位", 3号梯下端站第1限位 <- "输入_3号梯下端站第1限位", 3号梯下端站第2限位 <- "输入_3号梯下端站第2限位", 4号梯上端站第1限位 <- "输入_4号梯上端站第1限位", 4号梯上端站第2限位 <- "输入_4号梯上端站第2限位", 4号梯下端站第1限位 <- "输入_4号梯下端站第1限位", 4号梯下端站第2限位 <- "输入_4号梯下端站第2限位", 5号梯上端站第1限位 <- "输入_5号梯上端站第1限位", 5号梯上端站第2限位 <- "输入_5号梯上端站第2限位", 5号梯下端站第1限位 <- "输入_5号梯下端站第1限位", 5号梯下端站第2限位 <- "输入_5号梯下端站第2限位", 6号梯上端站第1限位 <- "输入_6号梯上端站第1限位", 6号梯上端站第2限位 <- "输入_6号梯上端站第2限位", 6号梯下端站第1限位 <- "输入_6号梯下端站第1限位", 6号梯下端站第2限位 <- "输入_6号梯下端站第2限位", 1号超重_1 <- "输出_1号梯满载指示", 2号超重_1 <- "输出_2号梯满载指示", 3号超重_1 <- "输出_3号梯满载指示", 4号超重_1 <- "输出_4号梯满载指示", 5号超重_1 <- "输出_5号梯满载指示", 6号超重_1 <- "输出_6号梯满载指示", 1号梯检修信号 <- "输入_1号梯检修信号", 2号梯检修信号 <- "输入_2号梯检修信号", 3号梯检修信号 <- "输入_3号梯检修信号", 4号梯检修信号 <- "输入_4号梯检修信号", 5号梯检修信号 <- "输入_5号梯检修信号", 6号梯检修信号 <- "输入_6号梯检修信号"

screen "1#电梯状态画面" 800x600
   Button "FB_Left_Square_1" at 391,451 size 20x20; TextOff 'Text'; PictureOff "FB_Left_Square_Released_256c"; PictureOn "FB_Left_Square_Pressed_256c"
      on Click: SetBit("输入_1号梯轿内关门按钮")
   Button "FB_Right_Square_1" at 371,451 size 20x20; TextOff 'Text'; PictureOff "FB_Right_Square_Released_256c_1"; PictureOn "FB_Right_Square_Pressed_256c"
      on Click: SetBit("输入_1号梯轿内关门按钮")
      Appearance <- "输入_1号梯轿内关门按钮"
   Button "FB_Left_Square" at 310,451 size 20x20; TextOff 'Text'; PictureOff "FB_Left_Square_Released_256c"; PictureOn "FB_Left_Square_Pressed_256c"
      on Click: SetBit("输入_1号梯轿内开门按钮")
   Button "FB_Right_Square" at 330,451 size 20x20; TextOff 'Text'; PictureOff "FB_Right_Square_Released_256c_1"; PictureOn "FB_Right_Square_Pressed_256c"
      on Click: SetBit("输入_1号梯轿内开门按钮")
      Appearance <- "输入_1号梯轿内开门按钮"
   TextField "文本域_1" at 385,8 size 281x43; Text '-- 1#电梯状态总览'
   TextField "文本域_3" at 68,13 size 292x31; Text '电 梯 监 控 系 统'
   Button "按钮_7" at 546,519 size 118x66; TextOff '电梯状态总览'
      on Click: ActivateScreen("电梯状态总览画面", 0)
   Button "按钮_8" at 669,519 size 111x66; TextOff '退出系统'
      on Click: StopRuntime(0)
   Group "Group_1" at 371,451 size 40x20; PictureOn "FB_Left_Square_Pressed_256c"; PictureOff "FB_Left_Square_Released_256c"
   Rectangle "矩形_193" at 167,126 size 4x18
      Appearance <- "输出_1号梯LEDi"
   Rectangle "矩形_194" at 167,148 size 4x18
      Appearance <- "输出_1号梯LEDj"
   Rectangle "矩形_195" at 180,124 size 18x4
      Appearance <- "输出_1号梯LEDa"
   Rectangle "矩形_196" at 177,128 size 4x18
      Appearance <- "输出_1号梯LEDf"
   Rectangle "矩形_197" at 180,145 size 18x4
      Appearance <- "输出_1号梯LEDg"
   Rectangle "矩形_198" at 177,149 size 4x18
      Appearance <- "输出_1号梯LEDe"
   Rectangle "矩形_199" at 180,167 size 18x4
      Appearance <- "输出_1号梯LEDd"
   Rectangle "矩形_200" at 197,127 size 4x18
      Appearance <- "输出_1号梯LEDb"
   Rectangle "矩形_201" at 197,149 size 4x18
      Appearance <- "输出_1号梯LEDc"
   Rectangle "矩形_237" at 75,311 size 44x21
      Appearance <- "输出_1号梯5层按钮指示灯"
   Rectangle "矩形_238" at 75,289 size 44x21
      Appearance <- "输出_1号梯6层按钮指示灯"
   Rectangle "矩形_239" at 75,267 size 44x21
      Appearance <- "输出_1号梯7层按钮指示灯"
   Rectangle "矩形_240" at 75,245 size 44x21
      Appearance <- "输出_1号梯8层按钮指示灯"
   Rectangle "矩形_241" at 75,223 size 44x21
      Appearance <- "输出_1号梯9层按钮指示灯"
   Rectangle "矩形_242" at 75,201 size 44x21
      Appearance <- "输出_1号梯10层按钮指示灯"
   Circle "圆_1" at 164,204 size 14x14
      Appearance <- "输出_10层下行呼梯按钮指示灯"
   Circle "圆_2" at 155,225 size 14x14
      Appearance <- "输出_9层上行呼梯按钮指示灯"
   Circle "圆_3" at 174,225 size 14x14
      Appearance <- "输出_9层下行呼梯按钮指示灯"
   Circle "圆_4" at 155,248 size 14x14
      Appearance <- "输出_8层上行呼梯按钮指示灯"
   Circle "圆_5" at 174,248 size 14x14
      Appearance <- "输出_8层下行呼梯按钮指示灯"
   Circle "圆_6" at 155,269 size 14x14
      Appearance <- "输出_7层上行呼梯按钮指示灯"
   Circle "圆_7" at 174,269 size 14x14
      Appearance <- "输出_7层下行呼梯按钮指示灯"
   Circle "圆_8" at 155,291 size 14x14
      Appearance <- "输出_6层上行呼梯按钮指示灯"
   Circle "圆_9" at 174,291 size 14x14
      Appearance <- "输出_6层下行呼梯按钮指示灯"
   Circle "圆_10" at 155,314 size 14x14
      Appearance <- "输出_5层上行呼梯按钮指示灯"
   Circle "圆_11" at 174,314 size 14x14
      Appearance <- "输出_5层下行呼梯按钮指示灯"
   Circle "圆_12" at 155,335 size 14x14
      Appearance <- "输出_4层上行呼梯按钮指示灯"
   Circle "圆_13" at 174,335 size 14x14
      Appearance <- "输出_4层下行呼梯按钮指示灯"
   Circle "圆_14" at 155,356 size 14x14
      Appearance <- "输出_3层上行呼梯按钮指示灯"
   Circle "圆_15" at 174,356 size 14x14
      Appearance <- "输出_3层下行呼梯按钮指示灯"
   Circle "圆_16" at 155,381 size 14x14
      Appearance <- "输出_2层上行呼梯按钮指示灯"
   Circle "圆_17" at 174,381 size 14x14
      Appearance <- "输出_2层下行呼梯按钮指示灯"
   Circle "圆_18" at 164,402 size 14x14
      Appearance <- "输出_1层上行呼梯按钮指示灯"
   TextField "文本域_41" at 77,432 size 48x19; Text '内呼'
   TextField "文本域_42" at 153,432 size 47x19; Text '外呼'
   Rectangle "矩形_233" at 75,399 size 44x21
      Appearance <- "输出_1号梯1层按钮指示灯"
   Rectangle "矩形_234" at 75,377 size 44x21
      Appearance <- "输出_1号梯2层按钮指示灯"
   Button "FB_Empty_Rectangular_1" at 83,401 size 29x18; TextOff 'Text'; PictureOff "FB_Empty_Rectangular_Released_256c"; PictureOn "FB_Empty_Rectangular_Pressed_256c"
      on Release: ResetBit("输入_1号梯轿内选层按钮1")
      on Press: SetBit("输入_1号梯轿内选层按钮1")
   Button "FB_Empty_Rectangular_2" at 83,379 size 29x18; TextOff 'Text'; PictureOff "FB_Empty_Rectangular_Released_256c"; PictureOn "FB_Empty_Rectangular_Pressed_256c"
      on Release: ResetBit("输入_1号梯轿内选层按钮2")
      on Press: SetBit("输入_1号梯轿内选层按钮2")
   Rectangle "矩形_235" at 75,355 size 44x21
      Appearance <- "输出_1号梯3层按钮指示灯"
   Button "FB_Empty_Rectangular_3" at 83,357 size 29x18; TextOff 'Text'; PictureOff "FB_Empty_Rectangular_Released_256c"; PictureOn "FB_Empty_Rectangular_Pressed_256c"
      on Release: ResetBit("输入_1号梯轿内选层按钮3")
      on Press: SetBit("输入_1号梯轿内选层按钮3")
   Rectangle "矩形_236" at 75,333 size 44x21
      Appearance <- "输出_1号梯4层按钮指示灯"
   Button "FB_Empty_Rectangular_4" at 83,335 size 29x18; TextOff 'Text'; PictureOff "FB_Empty_Rectangular_Released_256c"; PictureOn "FB_Empty_Rectangular_Pressed_256c"
      on Release: ResetBit("输入_1号梯轿内选层按钮4")
      on Press: SetBit("输入_1号梯轿内选层按钮4")
   Button "FB_Empty_Rectangular_5" at 83,313 size 29x18; TextOff 'Text'; PictureOff "FB_Empty_Rectangular_Released_256c"; PictureOn "FB_Empty_Rectangular_Pressed_256c"
      on Release: ResetBit("输入_1号梯轿内选层按钮5")
      on Press: SetBit("输入_1号梯轿内选层按钮5")
   Button "FB_Empty_Rectangular_6" at 83,291 size 29x18; TextOff 'Text'; PictureOff "FB_Empty_Rectangular_Released_256c"; PictureOn "FB_Empty_Rectangular_Pressed_256c"
      on Release: ResetBit("输入_1号梯轿内选层按钮6")
      on Press: SetBit("输入_1号梯轿内选层按钮6")
   Button "FB_Empty_Rectangular_7" at 83,269 size 29x18; TextOff 'Text'; PictureOff "FB_Empty_Rectangular_Released_256c"; PictureOn "FB_Empty_Rectangular_Pressed_256c"
      on Release: ResetBit("输入_1号梯轿内选层按钮7")
      on Press: SetBit("输入_1号梯轿内选层按钮7")
      Appearance <- "输出_1号梯7层按钮指示灯"
   Button "FB_Empty_Rectangular_8" at 83,247 size 29x18; TextOff 'Text'; PictureOff "FB_Empty_Rectangular_Released_256c"; PictureOn "FB_Empty_Rectangular_Pressed_256c"
      on Release: ResetBit("输入_1号梯轿内选层按钮8")
      on Press: SetBit("输入_1号梯轿内选层按钮8")
   Button "FB_Empty_Rectangular_9" at 83,225 size 29x18; TextOff 'Text'; PictureOff "FB_Empty_Rectangular_Released_256c"; PictureOn "FB_Empty_Rectangular_Pressed_256c"
      on Release: ResetBit("输入_1号梯轿内选层按钮9")
      on Press: SetBit("输入_1号梯轿内选层按钮9")
   Button "FB_Empty_Rectangular_10" at 83,203 size 29x18; TextOff 'Text'; PictureOff "FB_Empty_Rectangular_Released_256c"; PictureOn "FB_Empty_Rectangular_Pressed_256c"
      on Release: ResetBit("输入_1号梯轿内选层按钮10")
      on Press: SetBit("输入_1号梯轿内选层按钮10")
   TextField "文本域_14" at 90,399 size 14x19; Text '1'
   TextField "文本域_15" at 90,378 size 14x19; Text '2'
   TextField "文本域_16" at 90,355 size 14x19; Text '3'
   TextField "文本域_17" at 90,334 size 14x19; Text '4'
   TextField "文本域_18" at 90,312 size 14x19; Text '5'
   TextField "文本域_19" at 90,290 size 14x19; Text '6'
   TextField "文本域_20" at 90,268 size 14x19; Text '7'
   TextField "文本域_21" at 90,246 size 14x19; Text '8'
   TextField "文本域_22" at 90,224 size 14x19; Text '9'
   TextField "文本域_40" at 86,202 size 23x19; Text '10'
   Circle "圆_56" at 460,116 size 24x24
      Appearance <- "输出_1号梯满载指示"
   Circle "圆_57" at 570,116 size 24x24
      Appearance <- "输出_1号梯故障指示"
   Circle "圆_58" at 457,160 size 24x24
      Appearance <- "输出_1号梯照明指示"
   Circle "圆_60" at 568,162 size 24x24
      Appearance <- "输出_1号梯风扇指示"
   TextField "文本域_47" at 393,118 size 45x23; Text '超重'
   TextField "文本域_48" at 496,118 size 45x23; Text '满载'
   TextField "文本域_49" at 605,116 size 45x23; Text '故障'
   TextField "文本域_50" at 496,163 size 45x23; Text '照明'
   TextField "文本域_51" at 602,163 size 45x23; Text '风扇'
   Circle "圆_73" at 228,116 size 24x24
      Appearance <- "输入_自动运行信号"
   TextField "文本域_68" at 259,117 size 93x25; Text '自动运行'
   TextField "文本域_69" at 258,161 size 139x30; Text '电梯准备就绪'
   Circle "圆_19" at 228,160 size 24x24
      Appearance <- "输出_准备就绪信号"
   Group "Group" at 310,451 size 40x20; PictureOn "FB_Left_Square_Pressed_256c"; PictureOff "FB_Left_Square_Released_256c"
   Rectangle "矩形_1" at 93,114 size 6x34
      Appearance <- "输出_1号梯上行指示"
   Polygon "多边形_5" at 81,110 size 15x17
      Appearance <- "输出_1号梯上行指示"
   Polygon "多边形_6" at 96,110 size 14x17
      Appearance <- "输出_1号梯上行指示"
   Rectangle "矩形_73" at 93,149 size 6x34
      Appearance <- "输出_1号梯下行指示"
   Polygon "多边形_1" at 79,171 size 17x15
      Appearance <- "输出_1号梯下行指示"
   Polygon "多边形_2" at 96,171 size 17x15
      Appearance <- "输出_1号梯下行指示"
   Circle "圆_59" at 356,118 size 24x24
      Appearance <- "输出_1号梯满载指示"
   Circle "圆_83" at 620,279 size 16x16
      Appearance <- "输出_1号梯开门继电器"
   Circle "圆_86" at 620,295 size 16x16
      Appearance <- "输出_1号梯关门继电器"
   Circle "圆_129" at 620,229 size 16x16
      Appearance <- "输出_1号梯电机启动信号"
   Circle "圆_132" at 620,245 size 16x16
      Appearance <- "输出_1号梯上行接触器"
   Circle "圆_135" at 620,261 size 16x16
      Appearance <- "输出_1号梯下行接触器"
   TextField "文本域_97" at 521,280 size 92x15; Text '开门继电器'
   TextField "文本域_98" at 521,296 size 92x15; Text '关门继电器'
   TextField "文本域_104" at 521,261 size 92x15; Text '下行接触器'
   TextField "文本域_105" at 510,229 size 103x15; Text '电机启动信号'
   TextField "文本域_106" at 521,245 size 92x15; Text '上行接触器'
   Circle "圆_95" at 621,349 size 16x16
      Appearance <- "输出_1号梯1级减速制动"
   Circle "圆_98" at 621,364 size 16x16
      Appearance <- "输出_1号梯2级减速制动"
   Circle "圆_101" at 621,379 size 16x16
      Appearance <- "输出_1号梯3级减速制动"
   Circle "圆_104" at 621,318 size 16x16
      Appearance <- "输出_1号梯低速接触器"
   Circle "圆_107" at 621,333 size 16x16
      Appearance <- "输出_1号梯高速接触器"
   TextField "文本域_99" at 500,365 size 114x15; Text '二级制动接触器'
   TextField "文本域_100" at 500,381 size 114x15; Text '三级制动接触器'
   TextField "文本域_101" at 500,348 size 114x15; Text '一级制动接触器'
   TextField "文本域_102" at 500,316 size 114x15; Text '低速运行接触器'
   TextField "文本域_103" at 500,332 size 114x15; Text '高速运行接触器'
   Circle "圆_20" at 465,322 size 16x16
      Appearance <- "输入_1号梯检修信号"
   Circle "圆_21" at 465,338 size 16x16
      Appearance <- "输入_1号梯光幕信号"
   TextField "文本域_23" at 384,324 size 72x15; Text '检修开关'
   TextField "文本域_24" at 386,340 size 70x15; Text '光幕信号'
   Circle "圆_120" at 315,225 size 16x16
      Appearance <- "输入_1号梯10楼层门锁信号"
   Circle "圆_123" at 315,240 size 16x16
      Appearance <- "输入_1号梯9楼层门锁信号"
   Circle "圆_126" at 315,255 size 16x16
      Appearance <- "输入_1号梯8楼层门锁信号"
   Circle "圆_138" at 315,270 size 16x16
      Appearance <- "输入_1号梯7楼层门锁信号"
   Circle "圆_141" at 315,285 size 16x16
      Appearance <- "输入_1号梯6楼层门锁信号"
   Circle "圆_144" at 315,300 size 16x16
      Appearance <- "输入_1号梯5楼层门锁信号"
   Circle "圆_147" at 315,315 size 16x16
      Appearance <- "输入_1号梯4楼层门锁信号"
   Circle "圆_150" at 315,330 size 16x16
      Appearance <- "输入_1号梯3楼层门锁信号"
   Circle "圆_153" at 315,345 size 16x16
      Appearance <- "输入_1号梯2楼层门锁信号"
   Circle "圆_156" at 315,360 size 16x16
      Appearance <- "输入_1号梯1楼层门锁信号"
   Circle "圆_159" at 315,375 size 16x16
      Appearance <- "输入_1号梯轿厢门锁信号"
   TextField "文本域_76" at 219,227 size 91x15; Text '10层门锁信号'
   TextField "文本域_77" at 225,242 size 81x15; Text '9层门锁信号'
   TextField "文本域_78" at 225,256 size 81x15; Text '8层门锁信号'
   TextField "文本域_79" at 225,271 size 81x15; Text '7层门锁信号'
   TextField "文本域_80" at 225,286 size 81x15; Text '6层门锁信号'
   TextField "文本域_81" at 225,301 size 81x15; Text '5层门锁信号'
   TextField "文本域_83" at 225,316 size 81x15; Text '4层门锁信号'
   TextField "文本域_84" at 225,331 size 81x15; Text '3层门锁信号'
   TextField "文本域_85" at 225,346 size 81x15; Text '2层门锁信号'
   TextField "文本域_86" at 224,362 size 82x15; Text '1层门锁信号'
   TextField "文本域_87" at 225,376 size 81x15; Text '轿厢门锁信号'
   Circle "圆_162" at 465,227 size 16x16
      Appearance <- "输入_1号梯上端站第2限位"
   Circle "圆_165" at 465,242 size 16x16
      Appearance <- "输入_1号梯上端站第1限位"
   Circle "圆_168" at 465,257 size 16x16
      Appearance <- "输入_1号梯上平层信号"
   Circle "圆_171" at 465,272 size 16x16
      Appearance <- "输入_1号梯下平层信号"
   Circle "圆_174" at 465,287 size 16x16
      Appearance <- "输入_1号梯下端站第2限位"
   Circle "圆_177" at 465,302 size 16x16
      Appearance <- "输入_1号梯下端站第1限位"
   TextField "文本域_82" at 353,227 size 103x15; Text '上端站第二限位'
   TextField "文本域_88" at 352,243 size 104x15; Text '上端站第一限位'
   TextField "文本域_89" at 374,258 size 82x15; Text '上平层信号'
   TextField "文本域_90" at 374,273 size 82x15; Text '下平层信号'
   TextField "文本域_91" at 352,287 size 104x15; Text '下端站第二限位'
   TextField "文本域_92" at 352,303 size 104x15; Text '下端站第一限位'
   Circle "圆_22" at 466,358 size 16x16
      Appearance <- "输入_1号梯开门到位"
   Circle "圆_23" at 466,374 size 16x16
      Appearance <- "输入_1号梯关门到位"
   TextField "文本域_13" at 364,360 size 93x15; Text '开门到位信号'
   TextField "文本域_25" at 364,376 size 93x15; Text '关门到位信号'
   Clock "时钟_1" at 664,57 size 101x57
   DateTimeField "日期/时间域_1" at 491,71 size 184x28
   TextField "文本域_2" at 296,416 size 142x19; Text '1号电梯开关门状态'

